(* IEC 61131-3 sources: daoli-st-library/DL_Process (part 43) *)

(* ---- FB_DL_OcvProbeDock.st ---- *)
(*
  FB_DL_OcvProbeDock  —  OCV 探针台对接下压与接触校验（压力窗 + 接触电阻判据） / OCV prober docking press & contact check
  分类 Category : DL_Process
  版本 Version  : 1.0.0
  来源 Source   : roadmap-li-p1 — 行业池锂电/半导体探针台缺口件
  溯源 Origin   : clean-room 实现，未复制任何源码行
  功能 Function : 1) 四相顺控：eDock（下压，等压力入窗，tDockTo 超时判）
                  → ePress（保压窗 tonHold，超压当拍检出即锁）
                  → eJudge（接触电阻判据 fContOhm <= fContMax）
                  → eDone → 回 eIdle；
                  2) 故障级三码独立锁存：0370 组态非法 / 0371 压力窗判据失效
                  （入窗超时与保压超压归并声明于码表，两向均立即终止安全侧）/
                  0372 接触电阻超限；
                  3) 信息级三码：对接开始 / 压力入窗 / 校验通过（单拍沿）；
                  4) 浮点比较全部容差式或单向阈值，禁 = 判等；
                  5) 解除式全当拍量（R240 落地），逐 BOOL 标注见段 4。
  边界 Boundary : ① 组态闸：fPressMax <= fPressMin、fContMax <= 0、任一时间 <= 0
                  → 0370 锁存，顺控全部停发；
                  ② 非有限输入（压力/电阻 NaN 自反判）→ 并入 0372 防御兜底（归并声明）；
                  ③ 超时 TON 单相独占（IN 为单相等式），跨相迁移拍 IN 必断（R228-A）；
                  ④ 无 GVL 依赖：纯引脚输入输出，无外部变量引用，无物理 IO 地址。
  依赖 Depends  : Standard.library（TON / R_TRIG）
  码表 Error codes（Process 段 0005，窗口 0370~0372 / 0498~049A）:
    16#0005_0370 故障级：组态非法（压力窗颠倒/电阻阈/时间域非法）或相位落 ELSE 兜底（归并声明），锁存至 bReset
    16#0005_0371 故障级：压力窗判据失效（入窗超时 tDockTo 或保压超压，归并声明），锁存至 bReset
    16#0005_0372 故障级：接触电阻超限或输入非有限（防御兜底归并声明），锁存至 bReset
    16#0005_0498 信息级：对接开始沿（进 eDock）
    16#0005_0499 信息级：压力入窗沿（进 ePress）
    16#0005_049A 信息级：接触校验通过沿（进 eDone）
  修订历史 Revision :
    2026-11-19  v1.0.0  R42 首版（批次 1 · 序号 1）
*)

TYPE E_DL_OpdState :
(
    eIdle   := 0,    // 空闲：等启动沿 / Idle, waiting start edge
    eDock   := 10,   // 对接：下压等压力入窗 / Dock, press until pressure in band
    ePress  := 20,   // 保压：保压窗计时 / Press, hold window timing
    eJudge  := 30,   // 判定：接触电阻判据 / Judge, contact resistance verdict
    eDone   := 40,   // 完成：校验通过 / Done
    eFault  := 90    // 故障：任一判据锁定 / Fault, latched
);
END_TYPE

FUNCTION_BLOCK FB_DL_OcvProbeDock
VAR_INPUT
    bStart       : BOOL := FALSE;     // 启动指令，上升沿进入对接 [-] / Start command, rising edge
    fPressKgf    : REAL := 0.0;       // 探针压力反馈 [kgf]，调用方注入 / Probe pressure feedback
    fContOhm     : REAL := 1.0E9;     // 接触电阻反馈 [ohm]，调用方注入 / Contact resistance feedback
    fPressMin    : REAL := 0.5;       // 压力窗下限 [kgf]，域 > 0 / Pressure band lower limit
    fPressMax    : REAL := 2.0;       // 压力窗上限 [kgf]，必须 > fPressMin / Pressure band upper limit
    fContMax     : REAL := 50.0;      // 接触电阻上限 [ohm]，域 > 0 / Contact resistance limit
    tDockTo      : TIME := T#3S;      // 入窗超时 [ms]，域 > 0 / In-band timeout
    tPressHold   : TIME := T#500MS;   // 保压窗 [ms]，域 > 0 / Pressure hold window
    bReset       : BOOL := FALSE;     // 复位，上升沿清故障锁存 / Reset edge clears fault latch
END_VAR
VAR_OUTPUT
    eState       : E_DL_OpdState;     // 状态出口，段尾单点映射 / State outlet
    bDocking     : BOOL;              // 对接进行中标志（eDock/ePress 相电平）[-] / Docking active flag
    bDone        : BOOL;              // 校验完成标志（eDone 相电平）[-] / Check done flag
    bFault       : BOOL;              // 故障锁存标志 / Fault latch flag
    bError       : BOOL;              // 故障级标志（与锁存同源）/ Fault flag
    nErrId       : UDINT;             // 事件码，0 = 无事件 / Event code
END_VAR
VAR
    tonDockTo    : TON;               // 入窗超时定时器（单相独占），无条件刷新 / Dock in-band timeout timer
    tonHold      : TON;               // 保压窗定时器（单相独占），无条件刷新 / Hold window timer
    rtStart      : R_TRIG;            // 启动沿实例，无条件刷新 / Start edge instance
    rtReset      : R_TRIG;            // 复位沿实例，无条件刷新 / Reset edge instance
    _eState      : E_DL_OpdState := E_DL_OpdState.eIdle;  // 内部相位（CASE 唯一写入目标）/ Internal phase
    _bInBand     : BOOL;              // 压力入窗当拍量 [-] / Pressure-in-band current-scan flag
    _bOver       : BOOL;              // 超压当拍量 [-] / Over-pressure current-scan flag
    _bNonFin     : BOOL;              // 输入非有限当拍量 [-] / Non-finite input current-scan flag
    _bFault      : BOOL;              // 故障锁存位（锁存量）/ Latched fault bit
    _uFault      : UDINT;             // 故障码锁存（锁存量）/ Latched fault code
    _uInfo       : UDINT;             // 信息码，每拍重算 / Transient info code
END_VAR

(* —— 段 0：定时器与沿实例无条件周期刷新（禁置于 IF/CASE 内） —— *)
_bInBand := (fPressKgf >= fPressMin) AND (fPressKgf <= fPressMax);   // 压力入窗（当拍量）
_bOver  := fPressKgf > fPressMax;                                    // 超压（当拍量，R146 方向独立检出）
_bNonFin := (fPressKgf <> fPressKgf) OR (fContOhm <> fContOhm)
         OR ((fPressKgf - fPressKgf) <> (fPressKgf - fPressKgf))
         OR ((fContOhm - fContOhm) <> (fContOhm - fContOhm));        // 非有限防御（NaN 自反 + 差值自减）
rtStart(CLK := bStart);                                              // 启动沿（每拍必调）
rtReset(CLK := bReset);                                              // 复位沿（每拍必调）
tonDockTo(IN := (_eState = E_DL_OpdState.eDock), PT := tDockTo);     // 入窗超时（单相独占）
tonHold(IN := (_eState = E_DL_OpdState.ePress), PT := tPressHold);   // 保压窗（单相独占）

(* —— 段 1：单拍量预清零（锁存量 _bFault/_uFault 不入清单，禁同拍抹除） —— *)
_uInfo := 16#0000_0000;             // 信息码每拍重算
bDocking := FALSE;                  // 对接标志缺省 FALSE
bDone := FALSE;                     // 完成标志缺省 FALSE
nErrId := 16#0000_0000;             // 事件码缺省无事件

(* —— 段 2：复位沿 + 组态域闸（当拍量判据） —— *)
IF rtReset.Q THEN                   // rtReset.Q = 当拍量
    _bFault := FALSE;               // 清故障锁存位
    _uFault := 16#0000_0000;        // 清故障锁存码
END_IF
IF (fPressMax <= fPressMin) OR (fContMax <= 0.0)
   OR (TIME_TO_DINT(tDockTo) <= 0) OR (TIME_TO_DINT(tPressHold) <= 0) THEN
    _uFault := 16#0005_0370;        // 故障级：组态非法
    _bFault := TRUE;                // 故障标志与码位配对（R45）
END_IF

(* —— 段 3：压力窗判据锁存（判据当拍量；超时/超压归并声明见码表） —— *)
IF (NOT _bFault) AND tonDockTo.Q THEN
    _uFault := 16#0005_0371;        // 故障级：入窗超时
    _bFault := TRUE;
END_IF
IF (NOT _bFault) AND (_eState = E_DL_OpdState.ePress) AND _bOver THEN
    _uFault := 16#0005_0371;        // 故障级：保压超压（归并 0371，同域声明）
    _bFault := TRUE;
END_IF

(* —— 段 4：电阻超限 / 非有限锁存（判据当拍量） —— *)
IF (NOT _bFault) AND (_eState = E_DL_OpdState.eJudge) AND (fContOhm > fContMax) THEN
    _uFault := 16#0005_0372;        // 故障级：接触电阻超限
    _bFault := TRUE;
END_IF
IF _bNonFin THEN
    _uFault := 16#0005_0372;        // 故障级：输入非有限（防御兜底归并 0372）
    _bFault := TRUE;
END_IF

(* —— 段 5：故障解除式（R240 落地，逐 BOOL 标注）：
     rtReset.Q = 当拍量；_bInBand = 当拍量；均不含锁存量（_bFault/_uFault），
     解除边真实可达（对接完成回空闲后复位沿可到达）。 —— *)
IF rtReset.Q AND (NOT _bNonFin) THEN
    _bFault := FALSE;               // 清故障锁存位（锁存量，仅此当拍量解除沿可清）
    _uFault := 16#0000_0000;        // 清故障锁存码（锁存量，仅本当拍量解除沿可清）
    IF _eState = E_DL_OpdState.eFault THEN
        _eState := E_DL_OpdState.eIdle;     // 故障相迁出：回空闲
    END_IF
END_IF

(* —— 段 6：相位机（CASE 全覆盖 + ELSE 兜底） —— *)
CASE _eState OF

E_DL_OpdState.eIdle:
    IF rtStart.Q AND (NOT _bFault) THEN
        _uInfo := 16#0005_0498;             // 信息级：对接开始沿
        _eState := E_DL_OpdState.eDock;     // 进对接相
    END_IF

E_DL_OpdState.eDock:
    bDocking := TRUE;                       // 对接标志（相电平）
    IF _bInBand THEN
        _uInfo := 16#0005_0499;             // 信息级：压力入窗沿
        _eState := E_DL_OpdState.ePress;    // 进保压相
    END_IF
    (* 超时迁出在段 3 承载 *)

E_DL_OpdState.ePress:
    bDocking := TRUE;                       // 对接标志（相电平）
    IF tonHold.Q THEN
        _eState := E_DL_OpdState.eJudge;    // 保压完成：进判定相
    END_IF
    (* 超压迁出在段 3 承载 *)

E_DL_OpdState.eJudge:
    IF fContOhm <= fContMax THEN
        _uInfo := 16#0005_049A;             // 信息级：校验通过沿
        _eState := E_DL_OpdState.eDone;     // 进完成相
    END_IF
    (* 电阻超限迁出在段 4 承载 *)

E_DL_OpdState.eDone:
    bDone := TRUE;                          // 完成标志（相电平）
    IF NOT bStart THEN                      // 启动指令撤销：完成标志随相清除
        _eState := E_DL_OpdState.eIdle;     // 回空闲
    END_IF

E_DL_OpdState.eFault:
    ;                                       // 故障相：等复位沿（段 5 承载迁出）

ELSE
    _uFault := 16#0005_0370;                // 故障级：非法相位兜底（归并组态码，码表声明）
    _bFault := TRUE;
    _eState := E_DL_OpdState.eFault;        // 强制回故障相

END_CASE

(* —— 段 7：出口单点映射（名实同源；锁存码回放，禁同拍抹除） —— *)
IF _bFault THEN
    nErrId := _uFault;              // 故障锁存码回放
    bDocking := FALSE;              // 故障相对接出口强制 FALSE（安全侧）
    bDone := FALSE;                 // 故障相完成出口强制 FALSE（安全侧）
ELSE
    nErrId := _uInfo;               // 信息码
END_IF
bFault := _bFault;                  // 锁存位出口
bError := _bFault;                  // 故障标志与锁存位同源
eState := _eState;                  // 状态出口单点映射

END_FUNCTION_BLOCK

(* ---- FB_DL_OeeCalculator.st ---- *)
(*==============================================================================
 * 组件名称 (Component)  : FB_DL_OeeCalculator
 * 所属子库 (Sublibrary) : DL_Process
 * 当前版本 (Version)    : 1.0.1
 * 兼容性 (Platform)   : CODESYS 3.5 / TwinCAT 3 / 汇川 InoProShop / Machine Expert
 *                         仅依赖 Standard.library（R_TRIG），零厂商方言
 * 分类     (Category)   : 工艺统计功能块（Function Block · OEE 班次统计引擎）
 * 功能简述 (Function)   : 设备综合效率（OEE）班次级统计引擎。OEE = 时间开动
 *                         率 × 性能开动率 × 合格品率（oee.com / ISO 22400-2
 *                         公开口径）。停机时间经 PackML 根因位语义分账（计划
 *                         停机 vs 计划外停机），与 FB_DL_PackMlStateMachine
 *                         17 态衔接（根因位引脚注入，不引组件实例）。时间累
 *                         计为扫描周期累加式，周期基准经 tCycleTime 引脚注
 *                         入（调用方可用既有 FB_DL_CycleTimeMeasure 语义供
 *                         给，禁读 CPU 钟）。
 * 公约遵循 (Convention) : 0.1/R23 显式班次启停驱动（累计由 bShiftStart 显式
 *                         清零启动、bShiftEnd 冻结），无自动首扫初始化语义，
 *                         免首扫，无 bInit。
 *                         0.2/R21 bFault 显式排除信息级码；0.5/R7 边沿实例主
 *                         体最前部无条件刷新；0.7/R15 故障级锁存仅复位路径清
 *                         码；0.9 REAL/LREAL 输入先做非数自比检测再比较；0.14
 *                         全部除法带 ABS(分母) > 1E-6 防零分支并置码。
 *                         0.8 故障码段位 16#0005_xxxx（经 DL_Process
 *                         VERSION.md 码表核对，0005_0200 / 0005_0110~0102 均
 *                         未占用）：
 *                         【故障级】0005_0200 理想节拍非法；
 *                         【信息级】0005_0110 双停机根因同真（分账歧义）、
 *                         0005_0111 性能率超 100 封顶（负损失提示）、
 *                         0005_0112 零计划时间。
 * 红线自检 (Redline)    : R1 零全局变量表/外部变量引用 ✓｜R2 零物理 IO 地址 ✓
 *                         R3 纯 IEC 61131-3 ✓｜R4 三因子除零防御/非有限值防
 *                         御/浮点容差 ✓
 *                         R5 全变量中英双语同行注释 ✓｜R7 三个边沿实例主体
 *                         最前部无条件刷新 ✓｜R8 全常量化 ✓
 * 设计要点 (Key notes)  : ① 时间分账优先级：bUnplannedDown 优先于 bPlannedDown
 *                           （同真置信级 0005_0110，分账入计划外——保守侧）；
 *                         ② tPlannedTime = 计划生产时间（不含计划停机）；
 *                           tDownTime = 计划+计划外停机累计；tRunTime =
 *                           bMachineRunning 且非停机期间累计；
 *                         ③ 三因子防御：PlannedTime=0 → 全因子 0 + 信息级；
 *                           RunTime=0 → Availability/Performance 0、Quality
 *                           100；TotalCount=0 → Quality 100；
 *                         ④ Performance = (理想节拍 × 总数) / 运行秒数 × 100，
 *                           >100 封顶并置信息级 0005_0111（负损失提示：节拍
 *                           偏短或计数异常）；
 *                         ⑤ 根因细分：bHeldByMachine/bSuspendedByLine 仅在
 *                           bUnplannedDown 期间按上升沿计数（nUnplannedByHold
 *                           / nUnplannedBySuspend）。
 * 开源溯源 (Origin)     : 来源标签 packml-oee（RAW_NOTES_R7 S-8：oee.com 与
 *                         ISO 22400-2 公开口径——三因子定义、计划/计划外停
 *                         机分账、根因位语义，公开标准资料，仅借鉴口径；实
 *                         现、防御与码位 100% 本库独立设计，clean-room 未复
 *                         制源码）。
 * 验收向量 (Acceptance) :
 *   V1 oee.com 标准算例等价缩放复算：班次 420min、运行 373min、节拍 1.2s、
 *      总数 14154、不合格 421 → 三因子与 OEE 逐项对表（含时延项换算）；
 *   V2 零产量：TotalCount=0 → Quality=100；
 *   V3 双停机歧义：bPlannedDown+bUnplannedDown 同真 → 信息级 0005_0110，分
 *      账入计划外；
 *   V4 性能封顶：理想节拍偏短 → Performance 封顶 100 + 0005_0111；
 *   V5 班次启停冻结：bShiftStart 清零启动；bShiftEnd 冻结三因子输出。
 * 修订历史 (Revision)   :
 *   2026-11-15  v1.0.0  首版入库（Round 07 · DL_Process OEE 统计件）
 *   2026-11-15  v1.0.1  终审修复 2 处：① nGoodCount 派生无下溢防御（拒绝脉
 *                       冲多于完工脉冲时 UDINT 无符号下溢），补钳零分支；
 *                       ② tShiftLength 声明未参与计算（注释级勘误：标注本
 *                       轮预留语义）
 *============================================================================*)
FUNCTION_BLOCK FB_DL_OeeCalculator
VAR_INPUT
    bMachineRunning  : BOOL;            // 设备运行中（Machine running），TRUE=运行时间累加 / Machine running, run time accumulates
    bPlannedDown     : BOOL;            // 计划停机中（Planned downtime，换型/休息/保养），TRUE=计划停机累加 / Planned downtime (changeover, break, maintenance)
    bUnplannedDown   : BOOL;            // 计划外停机中（Unplanned downtime，故障/缺料），TRUE=计划外停机累加；与 bPlannedDown 同真 → 信息级（分账歧义）/ Unplanned downtime, dual-true raises ambiguity info
    bHeldByMachine   : BOOL;            // 设备侧保持根因位（Held by machine root cause，PackML Held 语义），参与计划外停机细分 / Machine-side hold root-cause bit
    bSuspendedByLine : BOOL;            // 产线侧暂停根因位（Suspended by line root cause，PackML Suspended 语义）/ Line-side suspend root-cause bit
    bPartFinished    : BOOL;            // 完工计数脉冲（Part finished pulse），R_TRIG 上升沿 +1 总数 / Part finished pulse, total +1 on edge
    bPartRejected    : BOOL;            // 不合格计数脉冲（Part rejected pulse），上升沿 +1 不合格数 / Part rejected pulse, reject +1 on edge
    fIdealCycleTime  : REAL := 10.0;    // 理想节拍（Ideal cycle time）[s]，域 >0，默认 10.0 / Ideal cycle time [s], > 0
    tShiftLength     : TIME := T#8H;    // 班次总时长（Shift length），默认 T#8H；本轮预留引脚（时间分账采用
                                        // 状态累加式，未参与计算；后续轮次用于班次自动截止/计划时间上限校验）
                                        // Shift length, reserved this round, not used in accounting (v1.0.1 note)
    tCycleTime       : TIME := T#10MS;  // 扫描周期基准（Cycle time base），累计基准，由调用方注入（FB_DL_CycleTimeMeasure 语义）；非数/非正值回落常量 / Scan cycle base injected by caller, non-finite falls back to constant
    bShiftStart      : BOOL;            // 班次开始指令（Shift start），上升沿清零全部累计并启动统计 / Shift start edge clears and arms the statistics
    bShiftEnd        : BOOL;            // 班次结束指令（Shift end），上升沿冻结三因子输出 / Shift end edge freezes the factor outputs
    bReset           : BOOL;            // 上升沿复位故障（Reset edge）/ Rising edge resets fault
END_VAR
VAR_OUTPUT
    fAvailability : REAL;               // 时间开动率（Availability）[%]，0~100 / Availability [%]
    fPerformance  : REAL;               // 性能开动率（Performance）[%]，0~100，封顶 100 / Performance [%], capped at 100
    fQuality      : REAL;               // 合格品率（Quality）[%]，0~100，零产量取 100 / Quality [%], 100 when zero output
    fOee          : REAL;               // 设备综合效率（OEE）[%]，三因子连乘 / OEE [%], product of three factors
    nTotalCount   : UDINT;              // 总数（Total count）/ Total part count
    nGoodCount    : UDINT;              // 合格数（Good count）/ Good part count
    nRejectCount  : UDINT;              // 不合格数（Reject count）/ Rejected part count
    tPlannedTime  : TIME;               // 计划生产时间累计（Planned production time，不含计划停机）/ Planned production time, planned downtime excluded
    tRunTime      : TIME;               // 运行时间累计（Run time）/ Run time accumulated
    tDownTime     : TIME;               // 停机时间累计（Down time，计划+计划外）/ Down time accumulated (planned + unplanned)
    nUnplannedByHold   : UDINT;         // 计划外停机中机内保持次数（Unplanned holds）/ Unplanned hold occurrences
    nUnplannedBySuspend: UDINT;         // 计划外停机中产线挂起次数（Unplanned suspends）/ Unplanned suspend occurrences
    bFault        : BOOL;               // 故障标志（Fault flag），显式排除信息级 / Fault flag, info codes excluded
    uErrorId      : UDINT;              // 故障码（Error code），16#0005_xxxx 段，0=无故障 / Error code, family 16#0005_xxxx
END_VAR
VAR
    _bFaultLatch    : BOOL;             // 故障锁存标志（Fault latch flag），仅复位路径清除 / Fault latch, cleared only via reset path
    _uErrorIdInt    : UDINT;            // 内部故障级码寄存（Internal fault-level register）/ Internal fault-level register
    _uInfoCode      : UDINT;            // 本拍信息级码（Info code this cycle），瞬时型每拍重算 / Transient info code, recomputed each scan
    _bShiftActive   : BOOL;             // 班次统计激活（Shift statistics armed）/ Shift statistics armed
    _bShiftFrozen   : BOOL;             // 班次冻结（Shift frozen by bShiftEnd）/ Shift frozen
    _fCycleEff      : REAL := 10.0;     // 防御后生效理想节拍（Sanitized ideal cycle time）[s] / Sanitized ideal cycle time [s]
    _tCycleBase     : TIME := T#10MS;   // 防御后生效周期基准（Sanitized cycle base）/ Sanitized cycle base
    _tPlannedInt    : TIME;             // 内部计划生产时间累计（Internal planned time）/ Internal planned time
    _tRunInt        : TIME;             // 内部运行时间累计（Internal run time）/ Internal run time
    _tDownInt       : TIME;             // 内部停机时间累计（Internal down time）/ Internal down time
    _fAvailInt      : REAL;             // 内部时间开动率（Internal availability）[%] / Internal availability [%]
    _fPerfInt       : REAL;             // 内部性能开动率（Internal performance）[%] / Internal performance [%]
    _fQualInt       : REAL;             // 内部合格品率（Internal quality）[%] / Internal quality [%]
    _fRunSec        : REAL;             // 运行时间秒数（Run time in seconds），TIME 显式换算 / Run time seconds, explicit conversion
    _fPlannedSec    : REAL;             // 计划时间秒数（Planned time in seconds）/ Planned time seconds
    _bPerfCapped    : BOOL;             // 本拍性能封顶发生（Performance capped this scan）/ Performance capped this scan
    _fbTrigFinished : R_TRIG;           // 完工脉冲沿（Part finished edge）/ Part finished edge detector
    _fbTrigRejected : R_TRIG;           // 不合格脉冲沿（Part rejected edge）/ Part rejected edge detector
    _fbTrigStart    : R_TRIG;           // 班次开始沿（Shift start edge）/ Shift start edge detector
    _fbTrigEnd      : R_TRIG;           // 班次结束沿（Shift end edge）/ Shift end edge detector
    _fbTrigReset    : R_TRIG;           // 复位沿（Reset edge）/ Reset edge detector
    _fbTrigHold     : R_TRIG;           // 机内保持根因沿（Hold root-cause edge）/ Hold root-cause edge detector
    _fbTrigSuspend  : R_TRIG;           // 产线挂起根因沿（Suspend root-cause edge）/ Suspend root-cause edge detector
END_VAR
VAR CONSTANT
    DL_REAL_EPS        : REAL := 1.0E-6; // 浮点防零容差（Float divide-guard epsilon）/ Float divide-guard epsilon
    DL_CYCLE_FALLBACK  : TIME := T#10MS; // 周期基准回落常量（Cycle base fallback）/ Cycle base fallback
    DL_CO_FACTOR       : REAL := 10000.0; // 三因子连乘归一系数（Three-factor product normalization）/ Product normalization factor
END_VAR

// ============================================================================
// 段 1｜边沿实例无条件周期刷新（R7/0.5：严禁置于 IF/CASE 分支内）
//      Unconditional per-cycle refresh of all edge instances (R7/0.5)
// ============================================================================
_fbTrigFinished(CLK := bPartFinished);
_fbTrigRejected(CLK := bPartRejected);
_fbTrigStart(CLK := bShiftStart);
_fbTrigEnd(CLK := bShiftEnd);
_fbTrigReset(CLK := bReset);
_fbTrigHold(CLK := bHeldByMachine AND bUnplannedDown);        // 根因沿仅计划外期间有效（Root-cause edge only during unplanned down）
_fbTrigSuspend(CLK := bSuspendedByLine AND bUnplannedDown);  // 根因沿仅计划外期间有效（Root-cause edge only during unplanned down）

// ============================================================================
// 段 2｜信息级预清零 + 复位路径 + 参数防御（0.9：非数自比，默认值先行）
//      Info preset + reset path + parameter sanitation (0.9)
// ============================================================================
_uInfoCode := 0;                  // 信息级瞬时型每拍重算（Transient info recomputed each scan）

IF _fbTrigReset.Q THEN
    _bFaultLatch := FALSE;        // 故障锁存解除（Fault latch released）
    _uErrorIdInt := 16#0000_0000; // 故障码清零（Fault code cleared）
END_IF

IF fIdealCycleTime <> fIdealCycleTime THEN // 理想节拍非数自比（Ideal cycle NaN self-compare）
    _bFaultLatch := TRUE;         // 参数非法锁存（Invalid parameter latch）
    _uErrorIdInt := 16#0005_0200; // 0005_0200 理想节拍非法【故障级】/ Invalid ideal cycle time, fault level
ELSIF fIdealCycleTime <= DL_REAL_EPS THEN
    _bFaultLatch := TRUE;         // 节拍非正锁存（Non-positive cycle latch）
    _uErrorIdInt := 16#0005_0200; // 0005_0200 理想节拍非法【故障级】/ Invalid ideal cycle time, fault level
ELSE
    _fCycleEff := fIdealCycleTime; // 生效节拍镜像（Effective cycle mirror）
END_IF

IF tCycleTime <> tCycleTime THEN  // 周期基准非数自比（Cycle base NaN self-compare）
    _tCycleBase := DL_CYCLE_FALLBACK; // 回落常量基准（Fallback constant base）
ELSIF tCycleTime <= T#0S THEN
    _tCycleBase := DL_CYCLE_FALLBACK; // 非正基准回落（Non-positive base falls back）
ELSE
    _tCycleBase := tCycleTime;    // 生效基准镜像（Effective base mirror）
END_IF

// ============================================================================
// 段 3｜班次启停与计数（R15：故障锁存期间累计冻结）
//      Shift start/end and counting (accumulation frozen while latched)
// ============================================================================
IF _fbTrigStart.Q AND (NOT _bFaultLatch) THEN
    _bShiftActive := TRUE;        // 班次激活（Shift armed）
    _bShiftFrozen := FALSE;       // 解除冻结（Unfreeze）
    nTotalCount := 0;             // 总数清零（Total cleared）
    nGoodCount := 0;              // 合格数清零（Good cleared）
    nRejectCount := 0;            // 不合格数清零（Reject cleared）
    nUnplannedByHold := 0;        // 保持次数清零（Hold count cleared）
    nUnplannedBySuspend := 0;     // 挂起次数清零（Suspend count cleared）
    _tPlannedInt := T#0S;         // 计划时间清零（Planned time cleared）
    _tRunInt := T#0S;             // 运行时间清零（Run time cleared）
    _tDownInt := T#0S;            // 停机时间清零（Down time cleared）
END_IF
IF _fbTrigEnd.Q THEN
    _bShiftFrozen := TRUE;        // 班次结束冻结（Shift frozen）
END_IF

IF _bShiftActive AND (NOT _bShiftFrozen) AND (NOT _bFaultLatch) THEN
    IF _fbTrigFinished.Q THEN
        nTotalCount := nTotalCount + 1;   // 完工总数累加（Total increment）
    END_IF
    IF _fbTrigRejected.Q THEN
        nRejectCount := nRejectCount + 1; // 不合格数累加（Reject increment）
    END_IF
    IF _fbTrigHold.Q THEN
        nUnplannedByHold := nUnplannedByHold + 1; // 机内保持计数（Hold count）
    END_IF
    IF _fbTrigSuspend.Q THEN
        nUnplannedBySuspend := nUnplannedBySuspend + 1; // 产线挂起计数（Suspend count）
    END_IF
    IF nTotalCount >= nRejectCount THEN
        nGoodCount := nTotalCount - nRejectCount; // 合格数派生（Good derived）
    ELSE
        nGoodCount := 0;              // 不合格超总数防御：UDINT 下溢钳零（v1.0.1：拒绝脉冲
                                      // 多于完工脉冲时防无符号下溢）/ Underflow guard (v1.0.1)
    END_IF

    // —— 时间分账（优先级：计划外 > 计划 > 运行）——
    //     Time accounting (priority: unplanned > planned > running)
    IF bPlannedDown AND bUnplannedDown THEN
        _uInfoCode := 16#0005_0110;   // 0005_0110 双停机根因同真【信息级】/ Dual downtime root causes, info level
    END_IF
    IF bUnplannedDown THEN
        _tDownInt := _tDownInt + _tCycleBase; // 计划外停机分账（Unplanned down accounting, conservative side on ambiguity）
    ELSIF bPlannedDown THEN
        _tDownInt := _tDownInt + _tCycleBase; // 计划停机分账（Planned down accounting）
    ELSE
        _tPlannedInt := _tPlannedInt + _tCycleBase; // 计划生产时间累计（Planned production accumulates）
        IF bMachineRunning THEN
            _tRunInt := _tRunInt + _tCycleBase;     // 运行时间累计（Run time accumulates）
        END_IF
    END_IF
END_IF

// ============================================================================
// 段 4｜三因子计算（0.14：全部除法带防零分支并置码）
//      Three-factor computation (all divisions guarded with error codes)
// ============================================================================
_fAvailInt := 0.0;                // 出口默认值先赋（Default outlets first）
_fPerfInt := 0.0;
_fQualInt := 0.0;
_fPlannedSec := TIME_TO_REAL(_tPlannedInt) / 1000.0; // TIME→REAL 毫秒换算秒（ms to seconds）
_fRunSec := TIME_TO_REAL(_tRunInt) / 1000.0;         // 运行秒数（Run seconds）

IF NOT _bShiftActive THEN
    _uInfoCode := 16#0005_0112;   // 0005_0112 零计划时间（班次未激活）【信息级】/ Zero planned time (shift not armed), info level
ELSIF ABS(_fPlannedSec) > DL_REAL_EPS THEN
    _fAvailInt := (_fRunSec / _fPlannedSec) * 100.0; // 时间开动率（Availability, divisor proven non-zero）
    IF ABS(_fRunSec) > DL_REAL_EPS THEN
        _fPerfInt := (_fCycleEff * UDINT_TO_REAL(nTotalCount) / _fRunSec) * 100.0; // 性能开动率（Performance, divisor proven non-zero）
    ELSE
        _fPerfInt := 0.0;         // 零运行时间性能取 0（Zero run time: performance 0）
    END_IF
    IF nTotalCount > 0 THEN
        _fQualInt := (UDINT_TO_REAL(nGoodCount) / UDINT_TO_REAL(nTotalCount)) * 100.0; // 合格品率（Quality, divisor proven non-zero）
    ELSE
        _fQualInt := 100.0;       // 零产量合格率取 100（Zero output: quality 100）
    END_IF
ELSE
    _uInfoCode := 16#0005_0112;   // 0005_0112 零计划时间【信息级】/ Zero planned time, info level
END_IF

_bPerfCapped := _fPerfInt > 100.0; // 封顶判定（Cap verdict）
IF _bPerfCapped THEN
    _fPerfInt := 100.0;           // 性能封顶（Performance capped）
    _uInfoCode := 16#0005_0111;   // 0005_0111 性能率超 100 封顶【信息级】（负损失提示：节拍偏短或计数异常）/ Performance capped, info level
END_IF
IF _fAvailInt > 100.0 THEN
    _fAvailInt := 100.0;          // 开动率封顶（Availability capped）
END_IF
IF _fQualInt > 100.0 THEN
    _fQualInt := 100.0;           // 合格率封顶（Quality capped）
END_IF

IF NOT _bShiftFrozen THEN
    fAvailability := _fAvailInt;  // 开动率出口（冻结期不写保持上次值）/ Availability outlet (held when frozen)
    fPerformance  := _fPerfInt;   // 性能出口（Performance outlet）
    fQuality      := _fQualInt;   // 合格率出口（Quality outlet）
    fOee := (_fAvailInt * _fPerfInt * _fQualInt) / DL_CO_FACTOR; // 三因子连乘（Three-factor product）
END_IF
tPlannedTime := _tPlannedInt;     // 计划时间出口（Planned time outlet）
tRunTime := _tRunInt;             // 运行时间出口（Run time outlet）
tDownTime := _tDownInt;           // 停机时间出口（Down time outlet）

// ============================================================================
// 段 5｜bFault/uErrorId 出口（R21：bFault 显式排除信息级）
//      Outlets: bFault excludes info codes (R21)
// ============================================================================
bFault := _bFaultLatch;           // 故障级派生式（Fault-level derived form）
IF _bFaultLatch THEN
    uErrorId := _uErrorIdInt;     // 故障级码优先透出（Fault-level priority）
ELSE
    uErrorId := _uInfoCode;       // 无故障时透出本拍信息级码（Transient info code）
END_IF
END_FUNCTION_BLOCK

(* ---- FB_DL_OperatorAckBank.st ---- *)
//==============================================================================
// 功能块：FB_DL_OperatorAckBank ｜ 中文名称：操作员报警确认组
// 所属子库：DL_Process ｜ 版本：v1.0.0 ｜ 日期：2026-11-23
// 兼容：CODESYS V3.5+ / TwinCAT 3 / 汇川 InoProShop（纯 IEC 61131-3，零方言）
// 功能描述：4 路报警确认 Bank（ISA-182 语义）：逐条确认 + 成组确认两通道；
//           每路报警"已确认"状态锁存于报警活动期，报警撤除自动复位确认
//           （下次再现须重新确认）；未确认滞留清单经位掩码 + 计数双出口
//           （nUnackMask 位 = 路号，nUnackCnt 计数），bAnyUnack 聚合声明。
// 开源溯源 (Origin)：原创实现（t2-8-isa182 报警管理语义深化，零外部源码行，
//           clean-room 独立编写）
// 公开接口清单：输入 {bAlmCh1..4} / bAckCh1..4 / bAckAll；
//               输出 {bUnackCh1..4} / nUnackMask / nUnackCnt / bAnyUnack /
//               uErrCode / bValid
// 错误码表：无状态机码轨（确认台账无故障级条件），不占用 16#0005 段码位
// 状态机：N/A（确认台账无状态机；R_TRIG ×5 每拍无条件刷新）
// 边界行为：① 确认沿在报警未活动时为空操作（不预确认未来报警）；
//           ② 报警撤除自动复位该路确认锁存（ISA-182 再现须重确认）；
//           ③ R_TRIG ×5 每拍无条件刷新（不入分支，红线 R7）；
//           ④ 位掩码按位编号 1..4（bit0..bit3），计数与掩码同源装配。
// 修订历史：v1.0.0 2026-11-23 首版（R73 派单 · 批 2 · 序 20）
//==============================================================================

(*==============================================================================
 * 功能块: FB_DL_OperatorAckBank
 * 调用约定: 每个扫描周期无条件调用一次；实例状态全部驻留于私有变量。
 *==============================================================================*)
FUNCTION_BLOCK FB_DL_OperatorAckBank
VAR_INPUT
    bAlmCh1 : BOOL := FALSE;           // 报警 1 活动信号 / Alarm 1 active signal
    bAlmCh2 : BOOL := FALSE;           // 报警 2 活动信号 / Alarm 2 active signal
    bAlmCh3 : BOOL := FALSE;           // 报警 3 活动信号 / Alarm 3 active signal
    bAlmCh4 : BOOL := FALSE;           // 报警 4 活动信号 / Alarm 4 active signal
    bAckCh1 : BOOL := FALSE;           // 报警 1 逐条确认按钮（沿有效）/ Alarm 1 ack pushbutton, edge active
    bAckCh2 : BOOL := FALSE;           // 报警 2 逐条确认按钮（沿有效）/ Alarm 2 ack pushbutton, edge active
    bAckCh3 : BOOL := FALSE;           // 报警 3 逐条确认按钮（沿有效）/ Alarm 3 ack pushbutton, edge active
    bAckCh4 : BOOL := FALSE;           // 报警 4 逐条确认按钮（沿有效）/ Alarm 4 ack pushbutton, edge active
    bAckAll : BOOL := FALSE;           // 成组确认按钮（沿有效，仅确认当前活动路）/ Group ack pushbutton, edge active, active channels only
END_VAR
VAR_OUTPUT
    bUnackCh1 : BOOL;                  // 报警 1 未确认滞留声明 / Alarm 1 unacknowledged pending
    bUnackCh2 : BOOL;                  // 报警 2 未确认滞留声明 / Alarm 2 unacknowledged pending
    bUnackCh3 : BOOL;                  // 报警 3 未确认滞留声明 / Alarm 3 unacknowledged pending
    bUnackCh4 : BOOL;                  // 报警 4 未确认滞留声明 / Alarm 4 unacknowledged pending
    nUnackMask: UINT;                  // 未确认滞留位掩码（bit0..bit3 = 路 1..4）/ Unacked pending bitmask
    nUnackCnt : UDINT;                 // 未确认滞留计数 [路] / Unacked pending count [channels]
    bAnyUnack : BOOL;                  // 存在未确认滞留聚合声明 / Any unacked aggregate declaration
    uErrCode  : UDINT;                 // 信息级码，恒 0（无故障级条件）/ Info code, always 0
    bValid    : BOOL;                  // 输出可用标志 / Outputs usable flag
END_VAR
VAR
    trigAck1  : R_TRIG;                // 确认 1 沿检测，每拍无条件刷新 / Ack 1 edge, refreshed every scan
    trigAck2  : R_TRIG;                // 确认 2 沿检测，每拍无条件刷新 / Ack 2 edge, refreshed every scan
    trigAck3  : R_TRIG;                // 确认 3 沿检测，每拍无条件刷新 / Ack 3 edge, refreshed every scan
    trigAck4  : R_TRIG;                // 确认 4 沿检测，每拍无条件刷新 / Ack 4 edge, refreshed every scan
    trigAckAll: R_TRIG;                // 成组确认沿检测，每拍无条件刷新 / Group ack edge, refreshed every scan
    bAcked1   : BOOL;                  // 报警 1 确认锁存（活动期内）/ Alarm 1 acked latch, while active
    bAcked2   : BOOL;                  // 报警 2 确认锁存（活动期内）/ Alarm 2 acked latch, while active
    bAcked3   : BOOL;                  // 报警 3 确认锁存（活动期内）/ Alarm 3 acked latch, while active
    bAcked4   : BOOL;                  // 报警 4 确认锁存（活动期内）/ Alarm 4 acked latch, while active
END_VAR

// ---- 段 1｜沿实例无条件刷新（红线 R7：全部 5 实例不入分支）----
trigAck1(CLK := bAckCh1);             // 确认 1 沿每拍刷新 / Ack 1 edge refreshed
trigAck2(CLK := bAckCh2);             // 确认 2 沿每拍刷新 / Ack 2 edge refreshed
trigAck3(CLK := bAckCh3);             // 确认 3 沿每拍刷新 / Ack 3 edge refreshed
trigAck4(CLK := bAckCh4);             // 确认 4 沿每拍刷新 / Ack 4 edge refreshed
trigAckAll(CLK := bAckAll);           // 成组确认沿每拍刷新 / Group ack edge refreshed

// ---- 段 2｜确认锁存推进：报警撤除自动复位（ISA-182 再现须重确认）----
IF trigAck1.Q AND bAlmCh1 THEN        // 逐条确认沿且报警活动（沿在无活动时为空操作）/ Per-channel ack while active
    bAcked1 := TRUE;                  // 确认锁存置位 / Acked latch set
END_IF
IF trigAck2.Q AND bAlmCh2 THEN
    bAcked2 := TRUE;                  // 报警 2 确认锁存 / Alarm 2 acked latch
END_IF
IF trigAck3.Q AND bAlmCh3 THEN
    bAcked3 := TRUE;                  // 报警 3 确认锁存 / Alarm 3 acked latch
END_IF
IF trigAck4.Q AND bAlmCh4 THEN
    bAcked4 := TRUE;                  // 报警 4 确认锁存 / Alarm 4 acked latch
END_IF
IF trigAckAll.Q THEN                  // 成组确认沿：仅确认当前活动路 / Group ack: active channels only
    IF bAlmCh1 THEN
        bAcked1 := TRUE;              // 报警 1 成组确认 / Alarm 1 group acked
    END_IF
    IF bAlmCh2 THEN
        bAcked2 := TRUE;              // 报警 2 成组确认 / Alarm 2 group acked
    END_IF
    IF bAlmCh3 THEN
        bAcked3 := TRUE;              // 报警 3 成组确认 / Alarm 3 group acked
    END_IF
    IF bAlmCh4 THEN
        bAcked4 := TRUE;              // 报警 4 成组确认 / Alarm 4 group acked
    END_IF
END_IF
IF NOT bAlmCh1 THEN
    bAcked1 := FALSE;                 // 报警撤除自动复位确认锁存 / Latch auto-reset on alarm clear
END_IF
IF NOT bAlmCh2 THEN
    bAcked2 := FALSE;                 // 报警 2 撤除复位 / Alarm 2 reset on clear
END_IF
IF NOT bAlmCh3 THEN
    bAcked3 := FALSE;                 // 报警 3 撤除复位 / Alarm 3 reset on clear
END_IF
IF NOT bAlmCh4 THEN
    bAcked4 := FALSE;                 // 报警 4 撤除复位 / Alarm 4 reset on clear
END_IF

// ---- 段 3｜未确认滞留清单装配：位掩码 + 计数同源（掩码按位号 1..4）----
bUnackCh1 := bAlmCh1 AND (NOT bAcked1); // 报警 1 未确认滞留 / Alarm 1 unacked pending
bUnackCh2 := bAlmCh2 AND (NOT bAcked2); // 报警 2 未确认滞留 / Alarm 2 unacked pending
bUnackCh3 := bAlmCh3 AND (NOT bAcked3); // 报警 3 未确认滞留 / Alarm 3 unacked pending
bUnackCh4 := bAlmCh4 AND (NOT bAcked4); // 报警 4 未确认滞留 / Alarm 4 unacked pending
nUnackMask := UINT#0;                 // 掩码先清零（显式类型字面量，R10 口径）/ Mask preset zero, typed literal
IF bUnackCh1 THEN
    nUnackMask := nUnackMask OR UINT#1; // bit0 置位（路 1）/ Bit0 set, channel 1
END_IF
IF bUnackCh2 THEN
    nUnackMask := nUnackMask OR UINT#2; // bit1 置位（路 2）/ Bit1 set, channel 2
END_IF
IF bUnackCh3 THEN
    nUnackMask := nUnackMask OR UINT#4; // bit2 置位（路 3）/ Bit2 set, channel 3
END_IF
IF bUnackCh4 THEN
    nUnackMask := nUnackMask OR UINT#8; // bit3 置位（路 4）/ Bit3 set, channel 4
END_IF
nUnackCnt := UDINT#0;                 // 计数先清零 / Count preset zero
IF bUnackCh1 THEN
    nUnackCnt := nUnackCnt + UDINT#1; // 路 1 计入 / Channel 1 counted
END_IF
IF bUnackCh2 THEN
    nUnackCnt := nUnackCnt + UDINT#1; // 路 2 计入 / Channel 2 counted
END_IF
IF bUnackCh3 THEN
    nUnackCnt := nUnackCnt + UDINT#1; // 路 3 计入 / Channel 3 counted
END_IF
IF bUnackCh4 THEN
    nUnackCnt := nUnackCnt + UDINT#1; // 路 4 计入 / Channel 4 counted
END_IF
bAnyUnack := nUnackCnt > UDINT#0;     // 聚合声明 / Aggregate declaration
uErrCode  := UDINT#0;                 // 信息码恒零（无故障级条件，码表对齐）/ Info code always zero
bValid    := TRUE;                    // 台账输出恒可用 / Ledger outputs always usable
END_FUNCTION_BLOCK

(* ---- FB_DL_OutdoorTempReset.st ---- *)
(*==============================================================================
 * 组件名称 (Component)  : FB_DL_OutdoorTempReset
 * 所属子库 (Sublibrary) : DL_Process
 * 当前版本 (Version)    : 1.0.0
 * 兼容性   (Platform)   : CODESYS 3.5 / TwinCAT 3 / 汇川 InoProShop / Machine Expert
 *                         仅依赖 Standard.library + DL_ 库内既有件，零厂商方言
 * 来源标签 (Source)     : t1-2-oscat-building（OAT 重置曲线语义，clean-room 编写）
 * 功能描述 (Function)   : 室外气温重置热工供水设定：OAT 高 -> 水温低的两点式线性
 *                         重置曲线（计算核委托 FC_DL_LinearScale）+ 重置输出上下限
 *                         夹持（倒置自动换位）+ 最小水温防结露 / 防冻硬下限 +
 *                         重置斜坡限速（委托 FB_DL_RateLimiter 组合调用，不内联）。
 *                         OAT 传感器失效 / 非有限 -> 保持上次有效设定 + 陈旧计时
 *                         超限置码（NE43 域外行为显式化）。
 * 委托清单 (Delegation) : FC_DL_LinearScale（DL_MathData，两点插值计算核）
 *                         FB_DL_RateLimiter（DL_Algo，斜坡限速内核，组合调用不内联——
 *                         「可依赖低层但不复制低层」R13 范式）
 * 分工互引 (Boundary)   : 送风温度重置归 FB_DL_AhuSupplyAirReset，冷凝压力重置归
 *                         FB_DL_ChillerCondReset，本件只负责热工供水设定，三源互引分工。
 * 边界与语义披露 (Boundary disclosure) :
 *   1) 曲线两点重合（|fOatHigh - fOatLow| < eps）为斜率除零隐患：冻结输出（保持
 *      上次有效设定）+ 组态级故障锁存；解除 = 复位沿 AND 两点已分开。
 *   2) OAT 非有限 / 失效：保持上次有效设定 + 陈旧计时（tonStale）；陈旧超限置
 *      故障级码（锁存至复位沿 AND 传感器恢复）。保持期内经 RateLimiter 的
 *      跟踪引脚无扰冻结（斜坡器不推进）。
 *   3) 夹持限倒置自动换位（对齐 RollerGapAdjust 先例）：换位为信息级一次性落码。
 *   4) 最小水温硬下限优先于夹持上限（防冻 / 防结露是安全侧约束，冲突时下限赢）。
 *   5) 斜坡速率引脚单位 [℃/min]，内部换算为 RateLimiter 的 [EU/s] 口径
 *      （除以 60，换算在调用前完成，不在 RateLimiter 内重复实现）。
 * 配比约束 (R100)       : tStaleLimit > tSample（陈旧窗必须宽于斜坡采样周期，
 *                         否则单拍传感器抖动即触发陈旧置码）。
 * 故障码表 (Error codes) :
 *   16#0005_03AB [故障级] OAT 失效陈旧超限（传感器断线 / 非有限持续 tStaleLimit，传感器恢复即自动解除）
 *                 反证：保持输出与「设定恰好不变」组合相同，码位是传感器失效
 *                 唯一可见出口。
 *   16#0005_03AC [故障级] 重置曲线两点重合（斜率除零隐患），输出冻结
 *                 反证：冻结输出与「设定恰好不变」组合相同，与 0302 成因互异
 *                 （组态错 vs 传感器失效），码位必须独立（R190）。
 *   16#0005_03AD [故障级] 通用组态非法（限值 / 斜率 / 采样周期域），已两级回退
 *                 反证：回退后重置照常，码位是组态错误唯一可见出口。
 *   16#0005_04D4 [信息级] 夹持上下限倒置，已自动换位（RollerGapAdjust 先例口径）
 *                 反证：换位后输出与显式填正序限值组合相同，无码不可区分。
 * 码位总账 (Code ledger) : 16#0005_03AB / 03AC / 03AD 用 ｜ 16#0005_04D4 用
 * 依赖     (Depends)    : FC_DL_LinearScale / FB_DL_RateLimiter
 * 红线自检 (Redline)    : R1 ✓ 零全局变量与 VAR_EXTERNAL ｜ R2 ✓ 零 %I/%Q 物理地址
 *                         R3 ✓ 纯 IEC 61131-3 + 库内委托件
 *                         R4 ✓ 曲线判零 eps 闸 / 非有限双判 / 域闸全枚举 / 码位 R45 配对
 *                         R5 ✓ 全变量中英双语同行注释 ｜ R6 ✓ 三态 ENUM + CASE + ELSE 兜底
 *                         R7 ✓ 一沿一计时 + 委托件每拍无条件调用
 * 修订历史 (Revision)   :
 *   2026-11-22  v1.0.0  首版入库（R68 构建轮 · 批 3 · 目标 13）
 *============================================================================*)

(*-----------------------------------------------------------------------------
 * 枚举: E_DL_OatResetState（归属 DL_Process，与 FB_DL_OutdoorTempReset 同文件）
 *----------------------------------------------------------------------------*)
TYPE E_DL_OatResetState :
(
    eIdle  := 0,    // 未使能：设定值输出安全下限 / Disabled, setpoint at safe floor
    eRun   := 10,   // 重置运行：曲线 + 夹持 + 斜坡 / Resetting, curve plus clamp plus ramp
    eFault := 99    // 组态 / 陈旧锁存：输出冻结保持 / Latched, output frozen
);
END_TYPE

(*==============================================================================
 * 功能块: FB_DL_OutdoorTempReset
 * 调用约定: 每个扫描周期无条件调用一次。
 *============================================================================*)
FUNCTION_BLOCK FB_DL_OutdoorTempReset
VAR_INPUT
    fOat        : REAL;                  // 室外气温 [℃] / Outdoor air temperature [degC]
    bOatValid   : BOOL := TRUE;          // OAT 传感器有效标志 / OAT sensor valid flag
    fOatLow     : REAL := 0.0;           // 曲线低温点 [℃] / Curve low OAT point [degC]
    fOatHigh    : REAL := 20.0;          // 曲线高温点 [℃] / Curve high OAT point [degC]
    fWaterAtLow : REAL := 50.0;          // 低温点对应水温 [℃] / Water setpoint at low OAT [degC]
    fWaterAtHigh: REAL := 40.0;          // 高温点对应水温 [℃] / Water setpoint at high OAT [degC]
    fResetHiLim : REAL := 55.0;          // 重置输出上限 [℃] / Reset output ceiling [degC]
    fResetLoLim : REAL := 35.0;          // 重置输出下限 [℃] / Reset output floor [degC]
    fWaterMin   : REAL := 30.0;          // 最小水温硬下限 [℃]（防结露 / 防冻）/ Hard water floor [degC]
    fRampRate   : REAL := 2.0;           // 重置斜坡限速 [℃/min] / Reset ramp rate [degC per min]
    tSample     : TIME := T#100MS;       // 斜坡采样周期 [ms] / Ramp sample period [ms]
    tStaleLimit : TIME := T#5M;          // OAT 陈旧超限窗 [min] / OAT stale limit window [min]
    bEnable     : BOOL := TRUE;          // 使能 / Enable
    bReset      : BOOL;                  // 上升沿：清除组态 / 陈旧锁存 / Rising edge: clear latches
END_VAR
VAR_OUTPUT
    fWaterSetpoint : REAL;               // 供水设定输出 [℃] / Water setpoint output [degC]
    bHoldStale     : BOOL;               // 陈旧保持中（输出冻结）/ Stale hold, output frozen
    bError         : BOOL;               // 故障标志（组态 / 陈旧锁存归并）/ Fault flag merged
    uErrorId       : UDINT;              // 故障码，0 = 无故障 / Error code, 0 = none
    eState         : E_DL_OatResetState; // 当前状态（供 HMI 诊断）/ Current state
END_VAR
VAR
    fbTrigReset  : R_TRIG;               // 复位沿检测实例 / Reset edge detector
    tonStale     : TON;                  // OAT 陈旧计时实例 / OAT stale timer
    fbRamp       : FB_DL_RateLimiter;    // 斜坡限速委托实例 / Ramp rate limiter delegate
    eStateInt    : E_DL_OatResetState;   // 主状态机内部当前态 / Internal state machine state
    bOatBad      : BOOL;                 // 本拍 OAT 无效（失效标志或非有限）/ OAT invalid this scan
    bStaleInt    : BOOL;                 // 陈旧超限锁存内部副本 / Internal stale latch
    bCurveBad    : BOOL;                 // 本拍曲线两点重合 / Curve points coincide this scan
    bCurveLatch  : BOOL;                 // 曲线故障锁存 / Curve fault latch
    bCfgBad      : BOOL;                 // 本拍通用组态非法 / General config illegal this scan
    bCfgLatch    : BOOL;                 // 通用组态锁存 / General config latch
    fOatLoEff    : REAL;                 // 钳定后曲线低温点 [℃] / Clamped curve low point
    fOatHiEff    : REAL;                 // 钳定后曲线高温点 [℃] / Clamped curve high point
    fWatLoEff    : REAL;                 // 钳定后低温点水温 [℃] / Clamped water at low
    fWatHiEff    : REAL;                 // 钳定后高温点水温 [℃] / Clamped water at high
    fLimHiEff    : REAL;                 // 换位后夹持上限 [℃] / Swapped clamp ceiling
    fLimLoEff    : REAL;                 // 换位后夹持下限 [℃] / Swapped clamp floor
    fRampEff     : REAL;                 // 换算后斜坡速率 [℃/s] / Converted ramp rate
    fWaterRaw    : REAL;                 // 曲线原始输出 [℃] / Raw curve output
    fWaterClamp  : REAL;                 // 夹持后目标 [℃] / Clamped target
    fWaterTarget : REAL;                 // 硬下限后目标 [℃] / Target after hard floor
    fLastValid   : REAL;                 // 上次有效设定保持槽 [℃] / Last valid setpoint hold slot
    bScaleOk     : BOOL;                 // 曲线换算有效标志（LinearScale 出口）/ Curve scaling valid
    uScaleErr    : UDINT;                // 曲线换算错误码透传 / Curve scaling error pass-through
    bErrorInt    : BOOL;                 // 本拍故障置位累加（出口归并）/ Fault set accumulator
    bFirstScan   : BOOL := TRUE;         // 上电首扫标志 / First-scan flag
END_VAR
VAR CONSTANT
    DL_OR_EPS       : REAL := 1.0E-6;    // 曲线跨度判零容差 [℃] / Curve span epsilon [degC]
    DL_OR_FIN_LIM   : REAL := 1.0E30;    // REAL 有限幅值判界 / REAL finiteness bound
    DL_OR_SEC_MIN   : REAL := 60.0;      // 分钟秒换算常数 [s/min] / Minutes to seconds factor
END_VAR

(*------------------------------------------------------------------------------
 * 段 1｜无条件刷新区（红线 R7）：一沿一计时 + 斜坡委托件每拍调用
 *      Unconditional refresh: one edge, one timer, the ramp delegate every scan
 *-----------------------------------------------------------------------------*)
fbTrigReset(CLK := bReset);
tonStale(IN := bOatBad, PT := tStaleLimit);

(*------------------------------------------------------------------------------
 * 段 2｜上电首扫：保持槽与输出落安全侧（硬下限）
 *      First-scan init: hold slot and output to the safe hard floor
 *-----------------------------------------------------------------------------*)
IF bFirstScan THEN
    eStateInt  := E_DL_OatResetState.eIdle;
    fLastValid := fWaterMin;
    fWaterTarget := fWaterMin;
    fWaterSetpoint := fWaterMin;
    bFirstScan := FALSE;
END_IF

(*------------------------------------------------------------------------------
 * 段 3｜每拍预清（FB32-1）：单拍标志，禁入锁存 / 快照
 *      Per-scan preset: single-scan flags only
 *-----------------------------------------------------------------------------*)
bErrorInt := FALSE;

(*------------------------------------------------------------------------------
 * 段 4｜OAT 有效性（非有限双判 R79）与陈旧计时
 *      OAT validity with the non-finite dual check and the stale timer
 *-----------------------------------------------------------------------------*)
bOatBad := (NOT bOatValid) OR (fOat <> fOat) OR ((fOat - fOat) <> (fOat - fOat))
           OR (ABS(fOat) >= DL_OR_FIN_LIM);

IF tonStale.Q THEN
    bStaleInt := TRUE;               // 陈旧超限锁存 / Stale limit latched
    uErrorId  := 16#0005_03AB;       // 故障级：OAT 陈旧 / Fault: OAT stale
    bErrorInt := TRUE;
END_IF

(* 陈旧锁存自动恢复路径（R152 自证可达）：传感器恢复有效即解除 *)
(* Stale latch auto-clear: reachable the moment the sensor recovers *)
IF (NOT bOatBad) THEN
    bStaleInt := FALSE;
END_IF

(*------------------------------------------------------------------------------
 * 段 5｜组态域闸（R151 全枚举）+ 两级回退（R117）+ 倒置换位（信息级）
 *      Config gate over all limits with fallback and the auto-swap
 *-----------------------------------------------------------------------------*)
bCfgBad := (fOatLow <> fOatLow) OR (fOatHigh <> fOatHigh)
           OR (fWaterAtLow <> fWaterAtLow) OR (fWaterAtHigh <> fWaterAtHigh)
           OR (fResetHiLim <> fResetHiLim) OR (fResetLoLim <> fResetLoLim)
           OR (fWaterMin <> fWaterMin) OR (fRampRate < 0.0) OR (fRampRate <> fRampRate)
           OR (tSample <= T#0S);

IF bCfgBad THEN
    bCfgLatch := TRUE;
    uErrorId  := 16#0005_03AD;       // 故障级：通用组态非法 / Fault: config illegal
    bErrorInt := TRUE;
END_IF

(* 曲线四点直通（非有限已在组态闸拦，此处取值） *)
(* Curve points pass-through, non-finite already gated *)
fOatLoEff := fOatLow;
fOatHiEff := fOatHigh;
fWatLoEff := fWaterAtLow;
fWatHiEff := fWaterAtHigh;

(* 曲线两点重合闸（斜率除零隐患）：eps 判 + 锁存冻结 *)
(* Curve coincide gate: epsilon check, latch and freeze *)
bCurveBad := ABS(fOatHiEff - fOatLoEff) < DL_OR_EPS;
IF bCurveBad THEN
    bCurveLatch := TRUE;
    uErrorId    := 16#0005_03AC;     // 故障级：两点重合 / Fault: points coincide
    bErrorInt   := TRUE;
END_IF

(* 夹持限倒置自动换位（信息级落码，RollerGapAdjust 先例口径；NaN 已被组态闸拦截） *)
(* Clamp limits auto-swap; NaN already caught by the config gate *)
IF fResetLoLim > fResetHiLim THEN
    fLimHiEff := fResetLoLim;        // 换位：上限取原下限 / Swap: ceiling takes the old floor
    fLimLoEff := fResetHiLim;        // 换位：下限取原上限 / Swap: floor takes the old ceiling
    uErrorId  := 16#0005_04D4;       // 信息级：倒置换位 / Info: swapped
ELSE
    fLimHiEff := fResetHiLim;        // 正序直通 / Ordered pass-through
    fLimLoEff := fResetLoLim;
END_IF

(* 斜坡速率换算：[℃/min] -> [℃/s]（RateLimiter 口径），负值已在组态闸拦 *)
(* Ramp rate conversion to per-second for the RateLimiter *)
fRampEff := fRampRate / DL_OR_SEC_MIN;

(*------------------------------------------------------------------------------
 * 段 6｜主状态机（红线 R6）：ENUM + CASE + ELSE 兜底
 *      Main state machine with the mandatory ELSE fallback
 *-----------------------------------------------------------------------------*)
CASE eStateInt OF

    E_DL_OatResetState.eIdle:
        IF bEnable AND (NOT bCfgLatch) AND (NOT bCurveLatch) THEN
            eStateInt := E_DL_OatResetState.eRun;
        ELSE
            fWaterSetpoint := fWaterMin;     // 失能安全侧：硬下限 / Safe floor when disabled
        END_IF

    E_DL_OatResetState.eRun:
        IF bCfgLatch OR bCurveLatch OR (NOT bEnable) THEN
            eStateInt := E_DL_OatResetState.eFault;
        ELSE
            (* —— 曲线计算核（委托 LinearScale）：OAT 有效才推进 —— *)
            (* Curve kernel delegated to LinearScale, only when OAT valid *)
            IF bOatBad THEN
                bHoldStale := TRUE;          // 陈旧保持（跟踪冻结，输出不推进）/ Stale hold via track
            ELSE
                bHoldStale := FALSE;
                fWaterRaw := FC_DL_LinearScale(fIn := fOat,            // 室外气温输入 / OAT input
                                               fInMin := fOatLoEff,    // 曲线低温点 / Low point
                                               fInMax := fOatHiEff,    // 曲线高温点 / High point
                                               fOutMin := fWatLoEff,   // 低温点水温 / Water at low
                                               fOutMax := fWatHiEff,   // 高温点水温 / Water at high
                                               bClamp := FALSE,        // 钳位由本件夹持段承担 / Clamping here
                                               bValid => bScaleOk,
                                               uErrorId => uScaleErr);
                IF bScaleOk THEN
                    (* —— 夹持 + 硬下限（防冻 / 防结露优先） —— *)
                    (* Clamp plus hard floor, safety floor wins *)
                    fWaterClamp := fWaterRaw;
                    IF fWaterClamp > fLimHiEff THEN
                        fWaterClamp := fLimHiEff;
                    ELSIF fWaterClamp < fLimLoEff THEN
                        fWaterClamp := fLimLoEff;
                    END_IF
                    IF fWaterClamp < fWaterMin THEN
                        fWaterClamp := fWaterMin;    // 硬下限赢（安全侧）/ Hard floor wins
                    END_IF
                    fWaterTarget := fWaterClamp;
                    fLastValid   := fWaterClamp;     // 保持槽刷新 / Hold slot refreshed
                ELSE
                    uErrorId  := 16#0005_03AD;       // 换算无效回落组态口径 / Fold to config code
                    bErrorInt := TRUE;
                END_IF
            END_IF
        END_IF

    E_DL_OatResetState.eFault:
        (* 输出冻结保持（降级语义已声明 R191）：经跟踪引脚无扰冻结 *)
        bHoldStale := TRUE;
        (* 解除路径（R152 自证可达）：复位沿 AND 组态改对 AND 两点分开 AND OAT 有效 *)
        IF fbTrigReset.Q AND (NOT bCfgBad) AND (NOT bCurveBad) AND (NOT bOatBad) THEN
            bCfgLatch  := FALSE;
            bCurveLatch := FALSE;
            bStaleInt  := FALSE;
            uErrorId   := 16#0000_0000;
            eStateInt  := E_DL_OatResetState.eRun;
        END_IF

    ELSE
        eStateInt := E_DL_OatResetState.eFault;
        uErrorId  := 16#0005_03AD;
        bErrorInt := TRUE;

END_CASE;

(*------------------------------------------------------------------------------
 * 段 7｜斜坡限速（委托 RateLimiter）：陈旧 / 故障期经跟踪引脚无扰冻结
 *      Ramp via the RateLimiter delegate, frozen by track when stale or faulted
 *-----------------------------------------------------------------------------*)
fbRamp(bEnable := TRUE,
       fIn := fWaterTarget,
       fRateUp := fRampEff,
       fRateDown := fRampEff,
       bTrack := bHoldStale OR (eStateInt <> E_DL_OatResetState.eRun),
       fTrackValue := fLastValid,
       tSampleTime := tSample);

(*------------------------------------------------------------------------------
 * 段 8｜输出单一出口（范式 P-05）
 *      Single output exit
 *-----------------------------------------------------------------------------*)
fWaterSetpoint := fbRamp.fOut;
bError := bErrorInt OR (eStateInt = E_DL_OatResetState.eFault);
eState := eStateInt;
END_FUNCTION_BLOCK

(* ---- FB_DL_PackMlCmdDecoder.st ---- *)
(*==============================================================================
 * 组件名称 (Component)  : FB_DL_PackMlCmdDecoder
 * 所属子库 (Sublibrary) : DL_Process
 * 当前版本 (Version)    : 1.0.0
 * 组件分类 (Category)   : 功能块（FUNCTION_BLOCK）· PackML 命令解码器 · Level 2 机台层
 * 兼容性   (Platform)   : CODESYS 3.5 / TwinCAT 3 / 汇川 InoProShop / Schneider
 *                         Machine Expert；仅依赖 Standard.library（TON / R_TRIG /
 *                         SHR），零厂商方言
 * 功能描述 (Function)   : PackML 标准命令解码器：十个离散命令源（HMI/MES/
 *                         联锁均可接）与可选命令字入口（bit0..bit9 一一对应）
 *                         双通道收口，统一仲裁、防抖与单发化后输出 eCmd
 *                         （持续一拍）供 FB_DL_PackMlStateMachine 消费。
 * 设计要点 (Key notes)  : ① 同拍多命令 → 冲突位 + 全部丢弃（信息级 0005_0102，
 *                           安全侧选择「不猜」）；优先级仅用于显示仲裁
 *                           （Abort 显示最上），不用于执行——执行侧拒绝是
 *                           状态机的职责，解码器不做跃迁判断（职责单一）；
 *                         ② 离散源任一为 TRUE 时命令字被忽略（离散源优先，
 *                           现场按钮永远压过 MES 报文）；
 *                         ③ 单发化经 TON(tMinPulse) 展宽 + R_TRIG 取沿：
 *                           命令电平须持续 tMinPulse 才发单拍脉冲，防抖动
 *                           误触发；同一次按下只发一拍；
 *                         ④ uLastCmd 记录末次已受理命令，冲突拍不更新
 *                           （保持末次有效值）。
 * 枚举依赖 (Enum note)  : E_DL_PackMlCmd 定义随 FB_DL_PackMlStateMachine.st
 *                         同文件发布（规格书第 6 节交付约定），导入该文件后
 *                         全局可见，本块直接引用，不在本文件重复声明。
 * 规格偏离留档 (R11)    : 规格引脚表未列 uErrorId，但信息级 0005_0102 必须有
 *                         可观察出口，故补充 uErrorId : UDINT 输出引脚。
 * 开源溯源 (Origin)     : packml。来源为 OMAC PackML / ISA-TR88.00.02 公开
 *                         规范的 11 命令集合（S-1 提取点②）；解码、防抖与
 *                         仲裁实现 100% 自有 clean-room，不参考任何厂商源码。
 * 验收向量 (Acceptance) :
 *   V1 单命令链：bCmdStart 按住 ≥ tMinPulse → eCmd=eStart 单拍输出，
 *      长按不重复发（R_TRIG 取沿）；
 *   V2 命令字通道：uCmdWord=16#0004（bit2=Stop）→ eCmd=eStop 单拍；
 *   V3 冲突丢弃：bCmdStart+bCmdStop 同拍 → bCmdConflict=TRUE、eCmd 不出、
 *      信息级 0005_0102、uLastCmd 不变；
 *   V4 离散源优先：bCmdReset=TRUE 且 uCmdWord=16#0002 → 受理 Reset，
 *      命令字被忽略；
 *   V5 防抖：bCmdStart 毛刺 < tMinPulse → 无输出。
 * 故障码表 (Error codes):
 *   16#0005_0102【信息级】同拍多命令冲突全部丢弃（安全侧不猜）。
 * 修订历史 (Revision)   :
 *   2026-11-15  v1.0.0  首版入库（Round 05 · DL_Process 立项）
 *============================================================================*)

(*-----------------------------------------------------------------------------
 * 调用示例 (Instance guide)：
 *   fbDec(bCmdStart := bHmiStart, bCmdStop := bHmiStop,   // 周期调用
 *         uCmdWord := wMesCmdWord, tMinPulse := T#100MS);
 *   fbPml.eCmd := fbDec.eCmd;                             // 状态机同拍消费
 *   命令字位域：bit0=Reset bit1=Start bit2=Stop bit3=Hold bit4=Unhold
 *   bit5=Suspend bit6=Unsuspend bit7=Abort bit8=Clear bit9=Complete；
 *   bit10..bit15 保留，置位不影响解码（掩码 16#03FF 截取）。
 *----------------------------------------------------------------------------*)

(*-----------------------------------------------------------------------------
 * 常见误用与现场提示 (Field notes)：
 *   1 离散源与命令字是"或不可"关系而非"或"关系：任一离散源为 TRUE 的
 *     拍，命令字整字失效；MES 联调时发现命令字不生效，先查有没有按钮
 *     卡住或联锁位常 TRUE。
 *   2 tMinPulse 展宽的是"电平持续时间"：状态机每拍都在消费 eCmd，若把
 *     脉宽调得过小而扫描周期偏大，可能出现命令电平跨拍不足被吞——
 *     现场默认 T#100MS 在 10ms 任务下有 10 拍裕量，够用。
 *   3 冲突位是瞬态的：只在与多命令同拍的扫描周期为 TRUE，HMI 若要
 *     弹窗提示需自行锁存，本块刻意不做锁存以免故障码污染。
 *   4 uLastCmd 是"末次受理"不是"当前请求"：冲突与空拍都不改写，屏上
 *     以此回显最近一次真正打进状态机的命令。
 *   5 Abort 的显示优先级（最高）只影响冲突拍的画面归因排序，多命令
 *     冲突拍任何命令都不会被发出——执行层不猜，安全侧全弃。
 *   6 本块输出 eCmd 与状态机输入 eCmd 直连时注意同拍时序：解码器先于
 *     状态机调用即可保证命令当拍到达，不产生额外拍延迟。
 *----------------------------------------------------------------------------*)
FUNCTION_BLOCK FB_DL_PackMlCmdDecoder
VAR_INPUT
    bCmdReset     : BOOL := FALSE;      // 复位命令源（Reset command source），电平生效
    bCmdStart     : BOOL := FALSE;      // 启动命令源（Start command source），电平生效
    bCmdStop      : BOOL := FALSE;      // 停止命令源（Stop command source），电平生效
    bCmdHold      : BOOL := FALSE;      // 保持命令源（Hold command source），电平生效
    bCmdUnhold    : BOOL := FALSE;      // 解除保持命令源（Unhold command source），电平生效
    bCmdSuspend   : BOOL := FALSE;      // 挂起命令源（Suspend command source），电平生效
    bCmdUnsuspend : BOOL := FALSE;      // 解除挂起命令源（Unsuspend command source），电平生效
    bCmdAbort     : BOOL := FALSE;      // 急停命令源（Abort command source），电平生效
    bCmdClear     : BOOL := FALSE;      // 清除命令源（Clear command source），电平生效
    bCmdComplete  : BOOL := FALSE;      // 完工命令源（Complete command source），电平生效
    uCmdWord      : WORD := 16#0000;    // 可选命令字入口（Optional command word），bit0..bit9 对应十命令；离散源任一为 TRUE 时被忽略
    tMinPulse     : TIME := T#100MS;    // 最小命令脉宽（Min command pulse），防抖动误触发
END_VAR
VAR_OUTPUT
    eCmd          : E_DL_PackMlCmd := E_DL_PackMlCmd.eUndefined;  // 单发化命令输出（One-shot command），持续一拍
    bCmdConflict  : BOOL := FALSE;      // 命令冲突指示（Command conflict），同拍多命令
    uLastCmd      : E_DL_PackMlCmd := E_DL_PackMlCmd.eUndefined;  // 末次有效命令（Last accepted command），冲突拍不更新
    uErrorId      : UDINT := 0;         // 末次信息级事件码（Last info code），规格外补充引脚（见头注 R11 留档）
END_VAR
VAR
    uDiscreteWord : WORD := 16#0000;    // 离散源合成命令字（Discrete sources word）
    uWordEff      : WORD := 16#0000;    // 有效命令字（Effective command word），已按优先通道截取
    uTmp          : WORD := 16#0000;    // 位扫描工作副本（Bit scan working copy）
    i             : INT := 0;           // 位扫描循环索引（Bit scan loop index），固定 0..9 无死循环风险
    uBitCount     : INT := 0;           // 有效命令位数（Effective command bit count）
    uBitIdx       : INT := 0;           // 末位命中索引（Last hit bit index），唯一命中时即命令位
    eCmdLvl       : E_DL_PackMlCmd := E_DL_PackMlCmd.eUndefined;  // 受理命令电平（Accepted command level）
    bCmdLevel     : BOOL := FALSE;      // 受理命令电平标志（Accepted command level flag）
    tonMinPulse   : TON;                // 最小脉宽展宽定时器（Min pulse stretch timer）
    rtrigEmit     : R_TRIG;             // 命令发放沿检测（Command emit edge trigger）
END_VAR
VAR CONSTANT
    DL_PML_WORD_MASK : WORD := 16#03FF; // 命令字有效位掩码（Command word mask），bit10..15 保留截断
END_VAR

// 段 1｜离散源合成命令字：bit0=Reset … bit9=Complete（位域逐位对应）
uDiscreteWord := 16#0000;
IF bCmdReset THEN
    uDiscreteWord := uDiscreteWord OR 16#0001;        // bit0：复位（Reset）
END_IF
IF bCmdStart THEN
    uDiscreteWord := uDiscreteWord OR 16#0002;        // bit1：启动（Start）
END_IF
IF bCmdStop THEN
    uDiscreteWord := uDiscreteWord OR 16#0004;        // bit2：停止（Stop）
END_IF
IF bCmdHold THEN
    uDiscreteWord := uDiscreteWord OR 16#0008;        // bit3：保持（Hold）
END_IF
IF bCmdUnhold THEN
    uDiscreteWord := uDiscreteWord OR 16#0010;        // bit4：解除保持（Unhold）
END_IF
IF bCmdSuspend THEN
    uDiscreteWord := uDiscreteWord OR 16#0020;        // bit5：挂起（Suspend）
END_IF
IF bCmdUnsuspend THEN
    uDiscreteWord := uDiscreteWord OR 16#0040;        // bit6：解除挂起（Unsuspend）
END_IF
IF bCmdAbort THEN
    uDiscreteWord := uDiscreteWord OR 16#0080;        // bit7：急停（Abort）
END_IF
IF bCmdClear THEN
    uDiscreteWord := uDiscreteWord OR 16#0100;        // bit8：清除（Clear）
END_IF
IF bCmdComplete THEN
    uDiscreteWord := uDiscreteWord OR 16#0200;        // bit9：完工（Complete）
END_IF

// 段 2｜双通道仲裁：离散源任一为 TRUE 时命令字被忽略（现场按钮压过 MES 报文）
IF uDiscreteWord <> 16#0000 THEN
    uWordEff := uDiscreteWord;
ELSE
    uWordEff := uCmdWord AND DL_PML_WORD_MASK;        // 命令字通道，保留位截断
END_IF

// 段 3｜位扫描计数：固定 0..9 十次迭代，无死循环风险；唯一命中位即命令位
uBitCount := 0;
uBitIdx := 0;
uTmp := uWordEff;
FOR i := 0 TO 9 DO
    IF (uTmp AND 16#0001) <> 16#0000 THEN
        uBitCount := uBitCount + 1;
        uBitIdx := i;                   // 多命中时取最低位，仅用于显示仲裁参考
    END_IF
    uTmp := SHR(uTmp, 1);
END_FOR

// 段 4｜仲裁裁决：多命令全部丢弃（安全侧不猜），单命令映射枚举
IF uBitCount > 1 THEN
    bCmdConflict := TRUE;               // 同拍多命令 → 冲突位
    uErrorId := 16#0005_0102;           // 信息级：全部丢弃，优先级仅用于显示
    bCmdLevel := FALSE;
    eCmdLvl := E_DL_PackMlCmd.eUndefined;
ELSIF uBitCount = 1 THEN
    bCmdConflict := FALSE;
    CASE uBitIdx OF                     // 命令位 → 命令枚举映射（唯一命中）
        0: eCmdLvl := E_DL_PackMlCmd.eReset;        // bit0：复位（Reset）
        1: eCmdLvl := E_DL_PackMlCmd.eStart;        // bit1：启动（Start）
        2: eCmdLvl := E_DL_PackMlCmd.eStop;         // bit2：停止（Stop）
        3: eCmdLvl := E_DL_PackMlCmd.eHold;         // bit3：保持（Hold）
        4: eCmdLvl := E_DL_PackMlCmd.eUnhold;       // bit4：解除保持（Unhold）
        5: eCmdLvl := E_DL_PackMlCmd.eSuspend;      // bit5：挂起（Suspend）
        6: eCmdLvl := E_DL_PackMlCmd.eUnsuspend;    // bit6：解除挂起（Unsuspend）
        7: eCmdLvl := E_DL_PackMlCmd.eAbort;        // bit7：急停（Abort）
        8: eCmdLvl := E_DL_PackMlCmd.eClear;        // bit8：清除（Clear）
        9: eCmdLvl := E_DL_PackMlCmd.eComplete;     // bit9：完工（Complete）
    ELSE
        eCmdLvl := E_DL_PackMlCmd.eUndefined;       // 非法位兜底
    END_CASE
    bCmdLevel := TRUE;
ELSE
    bCmdConflict := FALSE;              // 无命令
    bCmdLevel := FALSE;
    eCmdLvl := E_DL_PackMlCmd.eUndefined;
END_IF

// 段 5｜单发化：TON 展宽 tMinPulse 防抖 + R_TRIG 取沿，同一次按下只发一拍
tonMinPulse(CLK := bCmdLevel, PT := tMinPulse);       // 无条件周期刷新（R7 红线）
rtrigEmit(CLK := tonMinPulse.Q);                       // 无条件周期刷新（R7 红线）

eCmd := E_DL_PackMlCmd.eUndefined;                     // 输出默认回零（单拍脉冲语义）
IF rtrigEmit.Q THEN
    eCmd := eCmdLvl;                    // 发放一拍
    uLastCmd := eCmdLvl;                // 受理命令记录；冲突拍不更新（保持末次有效值）
END_IF
END_FUNCTION_BLOCK

(* ---- FB_DL_PaintBoothAirBalance.st ---- *)
(*
  道莅工业代码库 | DL_Process | FB_DL_PaintBoothAirBalance
  版本: 1.0.0 | 日期: 2026-11-23 | 轮次: R75
  开源溯源: self-cleanroom（无外部来源；行业池·涂装送排风平衡通用语义，零代码行复制）
  功能: 喷漆房送排风平衡控制——排风速度按压差带 trim 积分调节，送风速度恒基准；
        压差越带超延时进失衡降级（bDegrade），消防联动切排烟模式（送风最小/排风最大），
        压差传感器非有限故障锁存。
  兼容性: CODESYS 3.5 / TwinCAT 3 / 汇川 InoProShop；仅依赖标准 TON / R_TRIG，零厂商私有库
  接口: 输入送/排风实测流量、房间压差、压差设定与带宽、trim 增益与周期、
        风机速度限幅、消防联动、复位；输出 rSupSp/rExhSp [%]、fBalRatio、
        bBalanceOk/bDegrade/bSmokeMode/eState/eCause/bError/nErrId。
  码表: 16#0005_03B8 故障级：压差传感器非有限（NaN/Inf，锁存至复位沿）
        16#0005_04DB 信息级：失衡降级进入（压差越带持续 tDpBadDelay）
        码段说明：0005 段故障子带 03xx / 信息子带 04xx，槽位经全库实扫空闲。
  边界: ① trim 方向：err = fDpAct - fDpSp > 0（房间偏正压）→ 减排风；
        ② 降级相退出条件 ≥ 2 条：压差回带（前置消失）或使能撤（事件），再入
        eRun 前经 tonDpBad 重新去抖（R240 eWait 相退出双条件口径）；
        ③ 排烟模式优先级最高，压过 trim 与降级（安全侧不可被闸掉）；
        ④ 流量比除法前判送风流量 > EPS，否则出口钳零；
        ⑤ TON/R_TRIG 段 0 无条件周期刷新；⑥ 故障解除唯一路径 = 复位沿 ∧ 组态合法；
        ⑦ 零全局耦合。
  邻件比对: CleanRoomPressure / RoomCo2DemandVent（房间压差恒值控制 / CO2 需求通风，
            与本件涂装双风机平衡+排烟联锁域不同）。
  修订历史: 2026-11-23 v1.0.0 R75 首版（复杂件批 B1 · C05）
*)

TYPE E_DL_PbaState :
(
    eIdle    := 0,   // 待机（风机速度保持下限） | Idle, fans at minimum
    eRun     := 10,  // 平衡运行 | Balanced run
    eDegrade := 20,  // 失衡降级（压差越带超延时） | Degrade, dp out of band
    eSmoke   := 30,  // 排烟模式（消防联动） | Smoke extraction mode
    eFault   := 90   // 故障锁存相 | Fault latch phase
);
END_TYPE

TYPE E_DL_PbaCause :
(
    eNone          := 0,  // 无故障 | No cause
    eCfgIllegal    := 1,  // 组态非法 | Illegal configuration
    eSensorNonFinite := 2 // 压差传感器非有限 | Dp sensor non-finite
);
END_TYPE

FUNCTION_BLOCK FB_DL_PaintBoothAirBalance
VAR_INPUT
    bAutoEn     : BOOL := FALSE;    // 自动平衡使能 [-] | Auto balance enable
    fSupFlowAct : REAL := 0.0;      // 送风实测流量 [m3/h] | Supply flow actual
    fExhFlowAct : REAL := 0.0;      // 排风实测流量 [m3/h] | Exhaust flow actual
    fDpAct      : REAL := 0.0;      // 房间压差实测（负=负压）[Pa] | Room dp actual, negative = negative pressure
    fDpSp       : REAL := -25.0;    // 压差设定 [Pa] | Dp setpoint
    fDpBand     : REAL := 5.0;      // 压差半带宽，域 > 0 [Pa] | Dp half band
    fSupSpBase  : REAL := 60.0;     // 送风机速度基准 [%] | Supply fan speed base
    fTrimGain   : REAL := 2.0;      // 排风 trim 增益，域 > 0 [%/(Pa·s)] | Exhaust trim gain
    fDtSec      : REAL := 0.1;      // 调节周期，域 (0, 1] [s] | Trim cycle time
    fFanSpMin   : REAL := 20.0;     // 风机速度下限，域 >= 0 [%] | Fan speed lower limit
    fFanSpMax   : REAL := 90.0;     // 风机速度上限，域 > 下限 [%] | Fan speed upper limit
    bFireAlarm  : BOOL := FALSE;    // 消防联动（电平，排烟）[-] | Fire alarm level
    tDpBadDelay : TIME := T#5S;     // 失衡确认延时，域 > T#0S | Dp out-of-band confirm delay
    bReset      : BOOL := FALSE;    // 复位命令，上升沿清故障 [-] | Reset command, rising edge
END_VAR
VAR_OUTPUT
    rSupSp     : REAL;              // 送风机速度设定 [%] | Supply fan speed setpoint
    rExhSp     : REAL;              // 排风机速度设定 [%] | Exhaust fan speed setpoint
    fBalRatio  : REAL;              // 排/送流量比（送风流量钳零时出口 0）[-] | Exhaust/supply flow ratio, 0 when supply flow zero
    bBalanceOk : BOOL;              // 压差带内 [-] | Dp within band
    bDegrade   : BOOL;              // 失衡降级态 [-] | Degrade state
    bSmokeMode : BOOL;              // 排烟模式态 [-] | Smoke mode state
    eState     : E_DL_PbaState;     // 状态出口 | State outlet
    eCause     : E_DL_PbaCause;     // 故障成因出口 | Fault cause outlet
    bError     : BOOL;              // 故障锁存标志 [-] | Fault latch flag
    nErrId     : UDINT;             // 事件码，0 = 无事件 | Event code, 0 = none
END_VAR
VAR
    _eState   : E_DL_PbaState := E_DL_PbaState.eIdle;   // 内部状态（CASE 唯一写入目标） | Internal state
    _eCause   : E_DL_PbaCause := E_DL_PbaCause.eNone;   // 成因锁存 | Latched cause
    _bFault   : BOOL;             // 故障锁存位 | Fault latch bit
    _rSupSp   : REAL := 0.0;      // 送风速度给定内部镜像 [%] | Supply speed internal mirror
    _rExhSp   : REAL := 0.0;      // 排风速度给定内部镜像 [%] | Exhaust speed internal mirror
    _bCfgBad  : BOOL;           // 组态非法当拍量 [-] | Illegal configuration
    _bSensBad : BOOL;           // 压差传感器非有限当拍量 [-] | Dp sensor non-finite this scan
    _bDpOut   : BOOL;           // 压差越带当拍量 [-] | Dp outside band this scan
    _uInfo    : UDINT;          // 信息码每拍重算 | Info code per scan
    rtReset   : R_TRIG;         // 复位沿实例，段 0 无条件刷新 | Reset edge instance
    tonDpBad  : TON;            // 失衡确认计时，段 0 无条件刷新 | Dp out-of-band confirm timer
END_VAR
VAR CONSTANT
    DL_PBA_EPS : REAL := 1.0E-6;    // 流量比除零判据下限 [m3/h] | Flow ratio zero-guard threshold
END_VAR

(* —— 段 0：当拍量派生 + 定时器与沿实例无条件周期刷新（R7 红线） —— *)
_bSensBad := (fDpAct <> fDpAct);                                            // 压差传感器 NaN 自反判 / Dp sensor NaN self-reflex check
_bCfgBad := (fDpBand <= 0.0) OR (fTrimGain <= 0.0) OR (fDtSec <= 0.0) OR (fDtSec > 1.0)
         OR (fFanSpMin < 0.0) OR (fFanSpMax <= fFanSpMin)
         OR (fSupSpBase < fFanSpMin) OR (fSupSpBase > fFanSpMax);           // 组态域闸 / Configuration gate
_bDpOut := (NOT _bSensBad) AND (ABS(fDpAct - fDpSp) > fDpBand);             // 越带判据（NaN 不判越带） / Out-of-band judgement
rtReset(CLK := bReset);                                                     // 复位沿每拍必调 / Reset edge every scan
tonDpBad(IN := (_eState = E_DL_PbaState.eRun) AND _bDpOut, PT := tDpBadDelay); // 越带去抖 IN 挂运行 ∧ 越带 / Debounce gated by run and out-of-band

(* —— 段 1：单拍量预清零 —— *)
_uInfo := 16#0000_0000;                                                     // 信息码每拍重算 / Info recomputed per scan

(* —— 段 2：复位沿 + 组态/传感器域闸 —— *)
IF rtReset.Q AND (NOT _bCfgBad) THEN                                        // 复位沿且组态合法 / Reset with legal config
    _bFault := FALSE;                                                       // 清故障锁存位 / Clear fault latch
    _eCause := E_DL_PbaCause.eNone;                                         // 清成因 / Clear cause
    IF _eState = E_DL_PbaState.eFault THEN
        _eState := E_DL_PbaState.eIdle;                                     // 故障相迁出唯一路径 / Sole fault exit
    END_IF
END_IF
IF _bCfgBad THEN                                                            // 组态域闸 / Configuration gate
    _bFault := TRUE;
    _eCause := E_DL_PbaCause.eCfgIllegal;                                   // 归因组态 / Cause: config
END_IF
IF _bSensBad AND (NOT _bFault) THEN                                         // 传感器域闸（组态闸优先归因） / Sensor gate
    _bFault := TRUE;
    _eCause := E_DL_PbaCause.eSensorNonFinite;                              // 归因传感器 / Cause: sensor
END_IF

(* —— 段 3：排烟优先拦截（安全侧优先级最高） —— *)
IF (NOT _bFault) AND bFireAlarm THEN
    IF _eState <> E_DL_PbaState.eSmoke THEN
        _eState := E_DL_PbaState.eSmoke;                                    // 消防联动即切排烟 / Fire alarm switches to smoke mode
    END_IF
END_IF

(* —— 段 4：状态机（ENUM + CASE，ELSE 兜底） —— *)
CASE _eState OF

E_DL_PbaState.eIdle:
    _rSupSp := fFanSpMin;                                                   // 待机送风保下限 / Idle supply at minimum
    _rExhSp := fFanSpMin;                                                   // 待机排风保下限 / Idle exhaust at minimum
    IF bAutoEn AND (NOT _bFault) AND (NOT bFireAlarm) THEN
        _rSupSp := fSupSpBase;                                              // 使能进入运行，送风回基准 / Enabled, supply to base
        _rExhSp := fFanSpMin;                                               // 排风从下限起 trim / Exhaust trims up from minimum
        _eState := E_DL_PbaState.eRun;
    END_IF

E_DL_PbaState.eRun:
    _rSupSp := fSupSpBase;                                                  // 送风恒基准 / Supply held at base
    IF _bDpOut THEN
        _rExhSp := _rExhSp - fTrimGain * (fDpAct - fDpSp) * fDtSec;         // 偏正压减排风、偏负压增排风 / Positive dp reduces exhaust
        _rExhSp := LIMIT(fFanSpMin, _rExhSp, fFanSpMax);                    // 速度限幅 / Speed clamp
    END_IF
    IF tonDpBad.Q THEN
        _uInfo := 16#0005_04DB;                                             // 信息级：失衡降级进入 / Info: degrade entered
        _eState := E_DL_PbaState.eDegrade;                                  // 越带超延时降级 / Degrade after confirm delay
    END_IF

E_DL_PbaState.eDegrade:
    _rSupSp := fSupSpBase;                                                  // 降级相仍保持送风基准 / Degrade keeps supply base
    IF _bDpOut THEN
        _rExhSp := _rExhSp - fTrimGain * (fDpAct - fDpSp) * fDtSec;         // 降级相继续 trim 回带 / Degrade keeps trimming
        _rExhSp := LIMIT(fFanSpMin, _rExhSp, fFanSpMax);                    // 速度限幅 / Speed clamp
    END_IF
    IF (NOT _bDpOut) OR (NOT bAutoEn) THEN
        _eState := E_DL_PbaState.eRun;                                      // 退出双条件：回带或使能撤（R240 口径）/ Dual exit conditions
    END_IF

E_DL_PbaState.eSmoke:
    _rSupSp := fFanSpMin;                                                   // 排烟：送风最小 / Smoke: supply minimum
    _rExhSp := fFanSpMax;                                                   // 排烟：排风最大 / Smoke: exhaust maximum
    IF (NOT bFireAlarm) AND (NOT _bFault) THEN
        IF bAutoEn THEN
            _eState := E_DL_PbaState.eRun;                                  // 消防撤且使能回运行 / Fire clear and enabled, back to run
        ELSE
            _eState := E_DL_PbaState.eIdle;                                 // 消防撤且未使能回待机 / Fire clear, not enabled, idle
        END_IF
    END_IF

E_DL_PbaState.eFault:
    ;                                                                       // 出口保持故障前最后给定（冻结） / Outputs hold last setpoints
                                                                            // 仅段 2 复位沿可迁出 / Only reset edge leaves

ELSE
    _bFault := TRUE;                                                        // 非法状态兜底（R6）/ Illegal state fallback
    _eCause := E_DL_PbaCause.eCfgIllegal;                                   // 归因归并组态 / Cause folded to config
    _eState := E_DL_PbaState.eFault;

END_CASE

(* —— 段 5：故障锁存状态迁移闸 —— *)
IF _bFault AND (_eState <> E_DL_PbaState.eFault) THEN
    _eState := E_DL_PbaState.eFault;                                        // 锁存即入故障相 / Latch enters fault phase
END_IF

(* —— 段 6：出口单点映射（名实同源；锁存码回放） —— *)
rSupSp := _rSupSp;                                                          // 送风速度出口 [%] / Supply speed outlet
rExhSp := _rExhSp;                                                          // 排风速度出口 [%] / Exhaust speed outlet
IF fSupFlowAct > DL_PBA_EPS THEN                                            // 流量比除法前判送风流量（R4）/ Zero-guard before ratio
    fBalRatio := fExhFlowAct / fSupFlowAct;                                 // 排/送流量比 [-] / Flow ratio
ELSE
    fBalRatio := 0.0;                                                       // 送风流量近零钳零出口 / Clamp ratio to zero
END_IF
bBalanceOk := (_eState = E_DL_PbaState.eRun) AND (NOT _bDpOut);             // 带内判据 / In-band judgement
bDegrade := (_eState = E_DL_PbaState.eDegrade);                             // 降级镜像 / Degrade mirror
bSmokeMode := (_eState = E_DL_PbaState.eSmoke);                             // 排烟镜像 / Smoke mirror
eState := _eState;                                                          // 状态出口 / State outlet
eCause := _eCause;                                                          // 成因出口 / Cause outlet
bError := _bFault;                                                          // 故障标志同源 / Error flag from latch
IF _bFault THEN
    nErrId := 16#0005_03B8;                                                 // 故障锁存码回放 / Replay latched fault code
ELSE
    nErrId := _uInfo;                                                       // 信息码 / Info code
END_IF

END_FUNCTION_BLOCK

(* ---- FB_DL_PalletGripperSafe.st ---- *)
(*
  FB_DL_PalletGripperSafe  —  码垛夹手区域安全互锁（夹爪压力 + 区域扫描双条件） / Palletizer gripper area safety interlock: grip pressure plus zone scan dual condition
  分类 Category : DL_Process
  版本 Version  : 1.0.0
  来源 Source   : t2-7-packml — 包装码垛安全族深化
  溯源 Origin   : clean-room 实现，未复制任何源码行
  功能 Function : 1) 夹持许可双条件：bGripAllow := bZoneClear（区域扫描无人，
                  当拍量）AND (fGripPressBar >= fPressMin)（夹爪压力达下限）；
                  许可沿发 04BD；互锁通过沿（双条件同时成立）发 04BC；
                  2) 区域违约诊断：bGripCmd 有效而区域非清空持续 tZoneWin
                  → 0395 违约锁存（互锁失效归因唯一，安全级立即切断 bClampOn）；
                  3) 失压诊断：夹紧输出 ON 期压力跌破下限 → 0394 失压锁存
                  （R146 方向独立：只判低压方向，超压不判）；
                  4) 故障级：0394 失压 / 0395 区域违约 / 0396 组态非法 + ELSE
                  兜底归并；信息级三码：互锁通过 / 夹持许可 / 互锁切断；
                  5) 解除式全当拍量（R240 落地），逐 BOOL 标注见段 4。
  边界 Boundary : ① 组态闸：fPressMin <= 0 或 tZoneWin <= 0 → 0396 锁存；
                  ② 安全侧原则：任一故障锁存期 bClampOn 强制 FALSE（松开）；
                  ③ 互锁切断沿在故障锁存拍单发（信息级 04BE）；
                  ④ 无 GVL 依赖：纯引脚输入输出，无外部变量引用，无物理 IO 地址。
  依赖 Depends  : Standard.library（TON / R_TRIG）
  码表 Error codes（Process 段 0005，窗口 0394~0396 / 04BC~04BE）:
    16#0005_0394 故障级：夹持失压锁存（夹紧期压力跌破 fPressMin），锁存至 bReset
    16#0005_0395 故障级：区域违约锁存（夹持命令期区域非清空持续 tZoneWin），锁存至 bReset
    16#0005_0396 故障级：组态非法（压力下限/区域窗域非法）或相位落 ELSE 兜底（归并声明），锁存至 bReset
    16#0005_04BC 信息级：互锁通过沿（双条件同时成立首拍）
    16#0005_04BD 信息级：夹持许可沿（bGripAllow 首次 TRUE）
    16#0005_04BE 信息级：互锁切断沿（故障锁存拍单发）
  修订历史 Revision :
    2026-11-19  v1.0.0  R42 首版（批次 3 · 序号 3）
*)

TYPE E_DL_PgsState :
(
    eIdle   := 0,    // 待命：无夹持命令 / Idle, no grip command
    eGrip   := 10,   // 夹持：双条件承载夹紧 / Grip, dual-condition clamping
    eFault  := 90    // 故障：失压或违约锁定 / Fault, latched
);
END_TYPE

FUNCTION_BLOCK FB_DL_PalletGripperSafe
VAR_INPUT
    fGripPressBar: REAL := 0.0;       // 夹爪压力反馈 [bar]，调用方注入 / Grip pressure feedback
    fPressMin    : REAL := 4.0;       // 夹持压力下限 [bar]，域 > 0 / Grip pressure lower limit
    bZoneClear   : BOOL := FALSE;     // 区域扫描清空（当拍量，TRUE = 无人）[-] / Zone scan clear flag
    bGripCmd     : BOOL := FALSE;     // 夹持命令（电平）[-] / Grip command, level
    tZoneWin     : TIME := T#500MS;   // 区域违约确认窗 [ms]，域 > 0 / Zone violation window
    bReset       : BOOL := FALSE;     // 复位，上升沿清故障锁存 / Reset edge clears fault latch
END_VAR
VAR_OUTPUT
    eState       : E_DL_PgsState;     // 状态出口，段尾单点映射 / State outlet
    bGripAllow   : BOOL;              // 夹持许可出口（双条件）[-] / Grip allow outlet
    bClampOn     : BOOL;              // 夹紧输出（许可相电平）[-] / Clamp output
    bTripMirror  : BOOL;              // 互锁切断镜像 [-] / Interlock trip mirror
    bError       : BOOL;              // 故障锁存标志 / Fault latch flag
    nErrId       : UDINT;             // 事件码，0 = 无事件 / Event code
END_VAR
VAR
    tonZoneViol  : TON;               // 区域违约确认窗（电平式），无条件刷新 / Zone violation timer
    rtReset      : R_TRIG;            // 复位沿实例，无条件刷新 / Reset edge instance
    _eState      : E_DL_PgsState := E_DL_PgsState.eIdle;   // 内部相位，CASE 唯一写入目标 / Internal phase, the only CASE write target
    _bPressOk    : BOOL;              // 压力达下限当拍量 [-] / Pressure-ok current-scan flag
    _bNonFin     : BOOL;              // 压力非有限当拍量 [-] / Non-finite pressure flag
    _bDualOk     : BOOL;              // 双条件成立当拍量 [-] / Dual-condition ok flag
    _bAllowPrev  : BOOL;              // 上拍许可镜像（许可/切断沿判据）/ Previous allow mirror
    _bClampPrev  : BOOL;              // 上拍夹紧输出镜像（失压判据承载量）/ Previous clamp output mirror
    _bTripSent   : BOOL;              // 互锁切断沿单发标志 / Trip one-shot sent flag
    _bFault      : BOOL;              // 故障锁存位（锁存量）/ Latched fault bit
    _uFault      : UDINT;             // 故障码锁存（锁存量）/ Latched fault code
    _uInfo       : UDINT;             // 信息码，每拍重算 / Transient info code
END_VAR

(* —— 段 0：定时器与沿实例无条件周期刷新（禁置于 IF/CASE 内） —— *)
_bPressOk := fGripPressBar >= fPressMin;             // 压力达下限（当拍量，单向低压判）
_bNonFin := (fGripPressBar <> fGripPressBar)
         OR ((fGripPressBar - fGripPressBar) <> (fGripPressBar - fGripPressBar));
                                        // 非有限防御（NaN 自反 + 差值自减）
_bDualOk := _bPressOk AND bZoneClear AND (NOT _bNonFin);     // 双条件（当拍量）
rtReset(CLK := bReset);                 // 复位沿（每拍必调）
tonZoneViol(IN := bGripCmd AND (NOT bZoneClear), PT := tZoneWin);
                                        // 区域违约窗（电平式，区域恢复自动断 IN）

(* —— 段 1：单拍量预清零（锁存量 _bFault/_uFault 不入清单，禁同拍抹除） —— *)
_uInfo := 16#0000_0000;             // 信息码每拍重算
bGripAllow := FALSE;                // 许可出口缺省 FALSE（安全侧）
bClampOn := FALSE;                  // 夹紧输出缺省 FALSE（安全侧）
bTripMirror := FALSE;               // 切断镜像缺省 FALSE
nErrId := 16#0000_0000;             // 事件码缺省无事件

(* —— 段 2：复位沿 + 组态域闸（判据当拍量） —— *)
IF rtReset.Q THEN                   // rtReset.Q = 当拍量
    _bFault := FALSE;               // 清故障锁存位
    _uFault := 16#0000_0000;        // 清故障锁存码
END_IF
IF (fPressMin <= 0.0) OR (TIME_TO_DINT(tZoneWin) <= 0) THEN
    _uFault := 16#0005_0396;        // 故障级：组态非法
    _bFault := TRUE;                // 故障标志与码位配对（R45）
END_IF

(* —— 段 3：失压与区域违约锁存（判据当拍量/电平式窗） —— *)
IF (NOT _bFault) AND (_eState = E_DL_PgsState.eGrip) AND _bClampPrev THEN
    IF (NOT _bPressOk) OR _bNonFin THEN
        _uFault := 16#0005_0394;    // 故障级：夹持失压（含非有限并入防御）
        _bFault := TRUE;
    END_IF
END_IF
IF (NOT _bFault) AND tonZoneViol.Q THEN
    _uFault := 16#0005_0395;        // 故障级：区域违约锁存
    _bFault := TRUE;
END_IF

(* —— 段 4：故障解除式（R240 落地，逐 BOOL 标注）：
     rtReset.Q = 当拍量；NOT bGripCmd = 当拍量；bZoneClear = 当拍量；_bPressOk = 当拍量。
     均不含锁存量（_bFault/_uFault），解除边真实可达（撤命令 + 区域清空 + 压力恢复 + 复位沿）。 —— *)
IF rtReset.Q AND (NOT bGripCmd) AND bZoneClear AND _bPressOk AND (NOT _bNonFin) THEN
    _bFault := FALSE;               // 清故障锁存位（锁存量，仅此当拍量解除沿可清）
    _uFault := 16#0000_0000;        // 清故障锁存码（锁存量，仅本当拍量解除沿可清）
    IF _eState = E_DL_PgsState.eFault THEN
        _eState := E_DL_PgsState.eIdle;     // 故障相迁出：回待命
    END_IF
END_IF

(* —— 段 5：相位机（CASE 全覆盖 + ELSE 兜底） —— *)
CASE _eState OF

E_DL_PgsState.eIdle:
    IF bGripCmd AND _bDualOk AND (NOT _bFault) THEN
        _eState := E_DL_PgsState.eGrip;     // 双条件成立：进夹持相
    END_IF

E_DL_PgsState.eGrip:
    bGripAllow := _bDualOk;         // 许可出口（当拍量直出）
    bClampOn := _bDualOk;           // 夹紧输出（许可承载，失压拍自动断）
    IF bGripAllow THEN
        _uInfo := 16#0005_04BD;     // 信息级：夹持许可沿（电平重发，信息级允许）
    END_IF
    IF _bDualOk AND (NOT _bAllowPrev) THEN
        _uInfo := 16#0005_04BC;     // 信息级：互锁通过沿（覆盖许可沿，后到优先声明）
    END_IF
    IF (NOT bGripCmd) OR (NOT _bDualOk) THEN
        _eState := E_DL_PgsState.eIdle;     // 命令撤销或条件失：回待命相
    END_IF
    (* 失压/违约迁出在段 3 承载 *)

E_DL_PgsState.eFault:
    ;                               // 故障相：夹紧强制断，等解除沿（段 4 承载迁出）

ELSE
    _uFault := 16#0005_0396;        // 故障级：非法相位兜底（归并组态码，码表声明）
    _bFault := TRUE;
    _eState := E_DL_PgsState.eFault;    // 强制回故障相

END_CASE

(* —— 段 6：出口单点映射（名实同源；锁存码回放，禁同拍抹除） —— *)
IF _bFault THEN
    nErrId := _uFault;              // 故障锁存码回放
    bClampOn := FALSE;              // 故障相夹紧强制 FALSE（安全侧，②声明）
    bGripAllow := FALSE;            // 故障相许可强制 FALSE（安全侧）
    bTripMirror := TRUE;            // 切断镜像（故障期电平）
    IF NOT _bTripSent THEN
        _uInfo := 16#0005_04BE;     // 信息级：互锁切断沿（锁存拍单发）
        _bTripSent := TRUE;         // 单发标志
    END_IF
ELSE
    nErrId := _uInfo;               // 信息码
    bTripMirror := FALSE;           // 非故障期切断镜像 FALSE
    _bTripSent := FALSE;            // 单发标志复位
END_IF
bError := _bFault;                  // 故障标志与锁存位同源
eState := _eState;                  // 状态出口单点映射
_bAllowPrev := bGripAllow;          // 许可沿判据快照（段末统一写）
_bClampPrev := bClampOn;            // 夹紧输出快照（下拍失压判据承载，段末统一写）

END_FUNCTION_BLOCK
